(* IEC 61131-3 sources: daoli-st-library/DL_Motion (part 12) *)

(* ---- FB_DL_EdgeTrimTraverse.st ---- *)
(*==============================================================================
 * 组件名称 (Component)  : FB_DL_EdgeTrimTraverse
 * 所属子库 (Sublibrary) : DL_Motion
 * 当前版本 (Version)    : 1.0.0
 * 兼容性 (Platform)     : CODESYS 3.5 / TwinCAT 3 / 汇川 InoProShop（纯标准元素，零方言）
 * 功能描述 (Function)   : 修边刀架横动往复定位。启动后在行程两端之间往复，折返点按重叠量
 *                         外延，端点驻留可组态；停止请求只在段终点生效（半途硬切会在膜面
 *                         留刀痕）。行程过窄、速度出域判组态故障；目标越软包络在启动沿前
 *                         预检拒绝，一轴不动。不做刀压控制、不做随线速度联动、不做多段
 *                         变速。说明：既有 FB_DL_SoftLimitGuard 的契约绑定运动轴接口，
 *                         与本件的开环步进契约不同，故按同一语义内联预检，不做跨契约强转。
 * 溯源 (Origin)         : 道莅 clean-room 防御性实现
 * 本文件内含 (Contains) : TYPE E_DL_TraverseState / FUNCTION_BLOCK FB_DL_EdgeTrimTraverse
 * 依赖 (Depends)        : DL_Device/I_DL_StepperOpenLoop（只调用契约方法与属性）
 * 红线自检 (Redline)    : 无外部全局变量、无硬件地址直引 ｜ 全变量中英双语同行注释
 *                         行程宽度判零防除零 ｜ 重叠量与驻留出域双向钳制 ｜ 非有限用自反比较
 *                         驻留定时器与沿实例无条件周期刷新 ｜ 枚举显式赋值 ｜ CASE 含 ELSE
 * 错误码表 (Codes)      : 16#0004_033B 就绪（空闲/本拍无事件）
 *                         16#0004_033C 故障级 旋转轴/横动轴拒绝运动指令
 *                         16#0004_033D 故障级 组态非法（行程宽度 < 5 mm 或速度出域）
 *                         16#0004_033E 故障级 目标越软包络，启动沿前预检拒绝（一轴不动）
 *                         16#0004_033F 预留：本版不发码（下一轮区间起点，禁止回填）
 * 修订历史 (Revision)   : 2026-11-17  v1.0.0  首版入库 · R28 · 阶段三批 2
 * 验收向量 (Acceptance) : 正向 行程 0~300 mm、100 mm/s、重叠 5 mm、驻留 200 ms → 单程
 *                         约 3 s、端点重叠 5 mm、单程计数 +1
 *                         反向 行程改 0~3 mm（宽 3 mm < 5 mm）→ 16#0004_033D；重叠给
 *                         -50 mm → 钳 0 后照常运行；目标包络外延后越限 → 16#0004_033E
 *                         且一轴不动；轴拒绝指令 → 16#0004_033C
 *============================================================================*)

(*-----------------------------------------------------------------------------
 * 枚举: E_DL_TraverseState（归属本功能块，同文件发布，全库唯一定义）
 * 含义: 横动往复相位，每个成员在 CASE 中有且仅有一个标签。
 *----------------------------------------------------------------------------*)
TYPE E_DL_TraverseState :
(
    eIdle    := 0,    // 空闲：等启动沿与预检 / Idle, waiting for the start edge and the pre-check
    eRunMin  := 10,   // 向负端行进 / Travelling toward the minimum end
    eRunMax  := 20,   // 向正端行进 / Travelling toward the maximum end
    eDwell   := 30,   // 端点驻留计时 / Dwell timing at an end
    eStopped := 40,   // 段终点已停：等停止请求撤除 / Stopped at the segment end, waiting for the stop request to clear
    eFault   := 99    // 故障：锁存码保持，仅启动沿重启 / Fault, the latch code is held until a start edge
);
END_TYPE

FUNCTION_BLOCK FB_DL_EdgeTrimTraverse
VAR_INPUT
    bEnable       : BOOL := FALSE;        // 使能 / Enable
    bStart        : BOOL := FALSE;        // 启动，上升沿启动一次 / Start, the rising edge starts one cycle
    bStop         : BOOL := FALSE;        // 停止，电平请求，段终点生效 / Stop request, level input, effective at the segment end
    fPosMin_mm    : REAL := 0.0;          // 行程负端 [mm]，域 ±1000 / Negative travel end in millimetres, domain plus minus 1000
    fPosMax_mm    : REAL := 300.0;        // 行程正端 [mm]，须 Max − Min ≥ 5 / Positive travel end in millimetres, Max minus Min must reach 5
    fSpeed_mmS    : REAL := 100.0;        // 运行速度 [mm/s]，域 0.5~200 / Run speed in millimetres per second, domain 0.5 to 200
    fOverlap_mm   : REAL := 5.0;          // 端点重叠 [mm]，域 0~20 / End overlap in millimetres, domain 0 to 20
    tDwell        : TIME := T#200MS;      // 端点驻留 [ms]，域 0~5 s / End dwell, domain 0 to 5 s
END_VAR
VAR_IN_OUT
    iAxis         : I_DL_StepperOpenLoop; // 横动轴开环步进契约引用 [—] / Traverse axis open-loop stepper contract reference
END_VAR
VAR_OUTPUT
    fPosOut_mm    : REAL;                 // 当前横动位置 [mm] / Current traverse position in millimetres
    bAtMin        : BOOL;                 // 负端到位 / At the minimum end
    bAtMax        : BOOL;                 // 正端到位 / At the maximum end
    uTraverseCnt  : UDINT;                // 累计单程数 [次] / Accumulated single passes
    eState        : E_DL_TraverseState;   // 横动相位 [—] / Traverse phase
    eErr          : UDINT;                // 错误码，段位 16#0004_xxxx / Error code in segment 16#0004_xxxx
END_VAR
VAR
    _eState       : E_DL_TraverseState := E_DL_TraverseState.eIdle; // 当前相位 / Current phase
    _bInit        : BOOL := FALSE;        // 首扫标志，取非判定 / First-scan flag, tested negated
    _bRefOk       : BOOL;                 // 契约引用有效标志 / Contract reference valid flag
    _bCfgOk       : BOOL;                 // 组态合法标志 / Configuration valid flag
    _bIssueScan   : BOOL;                 // 派单当拍标志（本拍不判就绪） / Dispatch scan flag, readiness is not judged in this scan
    _bStopPending : BOOL;                 // 段终点停止挂起标志 / Stop pending at the segment end
    _bDirMax      : BOOL;                 // 下一段方向：TRUE = 向正端 / Next segment direction, TRUE for the positive end
    _bFaultLatch  : BOOL;                 // 故障锁存标志 / Fault latch flag
    _uLatchCode   : UDINT;                // 锁存码载体 / Latch code carrier
    _fTgtHigh     : REAL;                 // 正端折返目标（含重叠）[mm] / Positive turn target including overlap
    _fTgtLow      : REAL;                 // 负端折返目标（含重叠）[mm] / Negative turn target including overlap
    _fOverlapEff  : REAL := 0.0;          // 生效重叠量（钳制后）[mm] / Effective overlap after clamping
    _fSpeedEff    : REAL := 100.0;        // 生效速度（下限兜底）[mm/s] / Effective speed with a lower bound guard
    _fDist        : REAL;                 // 本段待走距离 [mm] / Pending distance of this segment
    _rtrigStart   : R_TRIG;               // 启动上升沿 / Rising edge of the start command
    _tonDwell     : TON;                  // 端点驻留计时 / End dwell timer
END_VAR
VAR CONSTANT
    DL_TRV_READY   : UDINT := 16#0004_033B;  // 就绪码 / Ready code
    DL_TRV_AXIS_BAD : UDINT := 16#0004_033C; // 故障级轴拒绝码 / Fault code for a rejected axis command
    DL_TRV_CFG_BAD : UDINT := 16#0004_033D;  // 故障级组态非法码 / Fault code for bad configuration
    DL_TRV_LIMIT   : UDINT := 16#0004_033E;  // 故障级预检拒绝码 / Fault code for a pre-check rejection
    DL_TRV_W_MIN   : REAL := 5.0;            // 行程最小宽度 [mm] / Minimum travel width in millimetres
    DL_TRV_POS_HI  : REAL := 1000.0;         // 行程端点绝对值上限 [mm] / Absolute bound of the travel ends
    DL_TRV_OVL_HI  : REAL := 20.0;           // 重叠量上限 [mm] / Overlap upper bound
    DL_TRV_SPD_LO  : REAL := 0.5;            // 速度下限 [mm/s] / Speed lower bound
    DL_TRV_SPD_HI  : REAL := 200.0;          // 速度上限 [mm/s] / Speed upper bound
    DL_TRV_AT_TOL  : REAL := 0.05;           // 端点到位容差 [mm] / End-point arrival tolerance
END_VAR

// 段 1｜输出与单拍标志预置
bAtMin := FALSE;                                    // 负端到位预清 / At-minimum flag pre-cleared
bAtMax := FALSE;                                    // 正端到位预清 / At-maximum flag pre-cleared
eErr := 0;                                          // 错误码预清 / Error code pre-cleared
_bIssueScan := FALSE;                               // 派单当拍标志预清 / Dispatch scan flag pre-cleared

// 段 2｜沿检测无条件周期刷新
_rtrigStart(CLK := bStart);                         // 启动沿 / Start edge

// 段 3｜驻留定时器无条件周期刷新（仅驻留相计时）
_tonDwell(IN := (_eState = E_DL_TraverseState.eDwell), PT := tDwell);

// 段 4｜首扫初始化（判据取非，R19）
IF NOT _bInit THEN
    _eState := E_DL_TraverseState.eIdle;            // 相位待机起步 / Phase starts idle
    _bInit := TRUE;                                 // 首扫只做一次 / The first scan runs once
END_IF

// 段 5｜引用与组态闸（行程宽度 < 5 mm 使往复退化为抖动）
_bRefOk := (iAxis <> 0);
_bCfgOk := _bRefOk
        AND NOT ((fPosMin_mm <> fPosMin_mm) OR ((fPosMin_mm - fPosMin_mm) <> (fPosMin_mm - fPosMin_mm)))
        AND NOT ((fPosMax_mm <> fPosMax_mm) OR ((fPosMax_mm - fPosMax_mm) <> (fPosMax_mm - fPosMax_mm)))
        AND ((fPosMax_mm - fPosMin_mm) >= DL_TRV_W_MIN)
        AND (ABS(fPosMin_mm) <= DL_TRV_POS_HI) AND (ABS(fPosMax_mm) <= DL_TRV_POS_HI)
        AND NOT ((fSpeed_mmS <> fSpeed_mmS) OR ((fSpeed_mmS - fSpeed_mmS) <> (fSpeed_mmS - fSpeed_mmS)))
        AND (fSpeed_mmS >= DL_TRV_SPD_LO) AND (fSpeed_mmS <= DL_TRV_SPD_HI)
        AND (tDwell >= T#0MS) AND (tDwell <= T#5S);
_fSpeedEff := LIMIT(DL_TRV_SPD_LO, fSpeed_mmS, DL_TRV_SPD_HI);          // 生效速度钳制 [mm/s] / Effective speed after clamping
_fOverlapEff := LIMIT(0.0, fOverlap_mm, DL_TRV_OVL_HI);                 // 重叠量钳制 [mm] / Overlap after clamping
_fTgtHigh := fPosMax_mm + _fOverlapEff;                                 // 正端折返目标（外延）[mm] / Positive turn target, extended
_fTgtLow := fPosMin_mm - _fOverlapEff;                                  // 负端折返目标（外延）[mm] / Negative turn target, extended

// 段 6｜位置回读与端点判据
IF _bRefOk THEN
    fPosOut_mm := iAxis.fPosition;                  // 当前横动位置 [mm] / Current traverse position
    bAtMax := ABS(fPosOut_mm - fTgtHigh) <= DL_TRV_AT_TOL;   // 正端到位判据 / At the positive end
    bAtMin := ABS(fPosOut_mm - fTgtLow) <= DL_TRV_AT_TOL;    // 负端到位判据 / At the negative end
ELSE
    fPosOut_mm := 0.0;                              // 引用无效：位置输出置 0 / Invalid reference, the position output is zeroed
END_IF

// 段 7｜失能闸
IF NOT bEnable THEN
    IF _bRefOk THEN
        iAxis.Stop();                               // 失能即受控停车 / Controlled stop on disable
    END_IF
    _eState := E_DL_TraverseState.eIdle;            // 相位回空闲 / Phase back to idle
    _bStopPending := FALSE;                         // 停止挂起清 / Stop pending cleared
    eErr := DL_TRV_READY;                           // 失能为正常停机 / Disable is a normal stop
END_IF

// 段 8｜横动往复状态机（ENUM + CASE + ELSE 兜底）
IF bEnable THEN
    CASE _eState OF

        E_DL_TraverseState.eIdle:                   // 空闲：等启动沿，先做组态与包络预检
            IF _rtrigStart.Q THEN
                _bFaultLatch := FALSE;              // 启动沿为锁存解除路径 / The start edge releases the latch
                _uLatchCode := 0;                   // 锁存码清 / Latch code cleared
                _bStopPending := FALSE;             // 停止挂起清 / Stop pending cleared
                IF NOT _bCfgOk THEN
                    eErr := DL_TRV_CFG_BAD;         // 故障级：组态非法 / Fault, bad configuration
                    _uLatchCode := DL_TRV_CFG_BAD;
                    _bFaultLatch := TRUE;
                    _eState := E_DL_TraverseState.eFault;
                ELSIF (ABS(_fTgtHigh) > DL_TRV_POS_HI) OR (ABS(_fTgtLow) > DL_TRV_POS_HI) THEN
                    eErr := DL_TRV_LIMIT;           // 故障级：重叠外延后越软包络，一轴不动 / Fault, the extended target leaves the envelope
                    _uLatchCode := DL_TRV_LIMIT;
                    _bFaultLatch := TRUE;
                    _eState := E_DL_TraverseState.eFault;
                ELSE
                    _bDirMax := TRUE;               // 首段向正端 / The first segment heads to the positive end
                    _eState := E_DL_TraverseState.eRunMax;
                END_IF
            ELSE
                IF NOT _bCfgOk THEN
                    eErr := DL_TRV_CFG_BAD;         // 故障级：组态非法（空闲期即报） / Fault, bad configuration reported while idle
                    _uLatchCode := DL_TRV_CFG_BAD;
                    _bFaultLatch := TRUE;
                    _eState := E_DL_TraverseState.eFault;
                END_IF
            END_IF

        E_DL_TraverseState.eRunMax:                 // 向正端行进：等轴就绪，停止请求挂起
            IF _bIssueScan THEN
                _bIssueScan := FALSE;               // 派单拍已过 / The dispatch scan has passed
            ELSIF (NOT _bStopPending) AND bStop THEN
                _bStopPending := TRUE;              // 停止请求挂起，段终点生效 / Stop pending, effective at the segment end
            ELSIF iAxis.bReady THEN
                uTraverseCnt := uTraverseCnt + 1;   // 单程计数 +1 [次] / Single-pass count incremented
                IF _bStopPending THEN
                    _eState := E_DL_TraverseState.eStopped;   // 段终点停车 / Stop at the segment end
                ELSE
                    _eState := E_DL_TraverseState.eDwell;     // 端点驻留 / Dwell at the end
                END_IF
            END_IF

        E_DL_TraverseState.eRunMin:                 // 向负端行进：等轴就绪，停止请求挂起
            IF _bIssueScan THEN
                _bIssueScan := FALSE;
            ELSIF (NOT _bStopPending) AND bStop THEN
                _bStopPending := TRUE;
            ELSIF iAxis.bReady THEN
                uTraverseCnt := uTraverseCnt + 1;   // 单程计数 +1 [次] / Single-pass count incremented
                IF _bStopPending THEN
                    _eState := E_DL_TraverseState.eStopped;
                ELSE
                    _eState := E_DL_TraverseState.eDwell;
                END_IF
            END_IF

        E_DL_TraverseState.eDwell:                  // 端点驻留：计时满后换向派单
            IF _tonDwell.Q THEN
                IF _bDirMax THEN
                    _bDirMax := FALSE;              // 换向：下一段向负端 / Reverse, the next segment heads to the negative end
                    _fDist := _fTgtLow - iAxis.fPosition;      // 待走距离 [mm] / Pending distance
                ELSE
                    _bDirMax := TRUE;               // 换向：下一段向正端 / Reverse, the next segment heads to the positive end
                    _fDist := _fTgtHigh - iAxis.fPosition;     // 待走距离 [mm] / Pending distance
                END_IF
                IF iAxis.MoveRelative(_fDist, _fSpeedEff) THEN
                    _bIssueScan := TRUE;            // 派单当拍不判就绪 / Readiness is not judged in the dispatch scan
                    IF _bDirMax THEN
                        _eState := E_DL_TraverseState.eRunMax;
                    ELSE
                        _eState := E_DL_TraverseState.eRunMin;
                    END_IF
                    eErr := DL_TRV_READY;           // 就绪码 / Ready code
                ELSE
                    eErr := DL_TRV_AXIS_BAD;        // 故障级：轴拒绝指令 / Fault, the axis rejected the command
                    _uLatchCode := DL_TRV_AXIS_BAD;
                    _bFaultLatch := TRUE;
                    _eState := E_DL_TraverseState.eFault;
                END_IF
            END_IF

        E_DL_TraverseState.eStopped:                // 段终点已停：停止请求撤除后回空闲
            IF NOT bStop THEN
                _bStopPending := FALSE;
                _eState := E_DL_TraverseState.eIdle;
            END_IF
            eErr := DL_TRV_READY;

        E_DL_TraverseState.eFault:                  // 故障：锁存码保持，仅新启动沿重启
            eErr := _uLatchCode;                    // 锁存码回放 / Replay the latch code
            IF _rtrigStart.Q THEN
                _bFaultLatch := FALSE;
                _uLatchCode := 0;
                _bStopPending := FALSE;
                eErr := DL_TRV_READY;
                _eState := E_DL_TraverseState.eIdle; // 回空闲需再给启动沿（下一拍） / A further start edge is required
            END_IF

        ELSE
            // 非法状态兜底（故障级）
            eErr := DL_TRV_CFG_BAD;                 // 故障级：非法相位 / Fault, illegal phase
            _uLatchCode := DL_TRV_CFG_BAD;
            _bFaultLatch := TRUE;
            _eState := E_DL_TraverseState.eFault;

    END_CASE
END_IF

eState := _eState;                                  // 相位出口镜像 / Phase mirrored to the output pin
END_FUNCTION_BLOCK

(* ---- FB_DL_ElectrodeRollDiameter.st ---- *)
// =====================================================================
// FB_DL_ElectrodeRollDiameter.st
// 极卷直径跟踪与换卷预警（卷径递推 + 低速保护 + 单调校核 + 换卷阈值预警）
// Electrode roll diameter tracking with change-over warning
// 所属子库: DL_Motion    版本: v1.0.0    兼容: CODESYS V3.5+ / TwinCAT 3 / 汇川 InoProShop
// 码位: 16#0004_035E ~ 16#0004_0362 (本件独占 5 槽, 勿复用)
// 溯源: 道莅 clean-room 防御性实现
//       来源组标签: lithium-battery, winding, coil-diameter, warning
// 修改记录: R30 初版 (ROUND_PLAN_R30 序 16)
// 分层声明: 卷径换算公式与 FC_DL_CoilDiameterCalc 口径一致（本件只加跟踪
//           与预警层, 不重写公式件）: D = v·k/(π·n), k = 1000 mm/m
// =====================================================================
FUNCTION_BLOCK FB_DL_ElectrodeRollDiameter
VAR_INPUT
    fLineSpd_mmin : REAL := 0.0;    // 线速度 0~300 m/min / Line speed [m/min]
    fRollRpm      : REAL := 0.0;    // 卷轴转速 0~3000 r/min / Roll speed [r/min]
    fPrevDia_mm   : REAL := 500.0;  // 上次卷径注入 0~2000 mm / Previous diameter injected [mm]
    fCoreDia_mm   : REAL := 76.0;   // 卷芯直径 0~2000 mm / Core diameter [mm]
    fThick_um     : REAL := 25.0;   // 层厚校核值 0~500 um / Layer thickness [um]
    fWarnDia_mm   : REAL := 120.0;  // 换卷预警径 0~2000 mm / Change warning diameter [mm]
END_VAR
VAR_OUTPUT
    fDia_mm     : REAL := 0.0;      // 当前卷径 / Current diameter [mm]
    bChangeWarn : BOOL := FALSE;    // 换卷预警 / Change-over warning
    bAtCore     : BOOL := FALSE;    // 卷径触及芯径 / At core flag
    eErr        : UDINT := 16#0004_035E;  // 错误码 / Error code
END_VAR
VAR
    rPi     : REAL := 3.14159265358979;   // 圆周率 / Pi constant
    fSpdMin : REAL := 1.0;          // 低速门限（线速度）m/min, 工程固定门限 / Min line speed gate
    fRpmMin : REAL := 5.0;          // 低速门限（转速）r/min, 工程固定门限 / Min roll speed gate
    fCalcDia: REAL := 0.0;          // 本拍换算卷径 / Calculated diameter this cycle [mm]
    fTolDia : REAL := 0.0;          // 单调校核容差（双倍层厚换算）/ Monotonic tolerance from thickness [mm]
    bCfgErr : BOOL := FALSE;        // 组态非法标记 / Configuration error flag
    bHoldErr: BOOL := FALSE;        // 递推保持标记（非有限或单调违反）/ Recursion hold flag
    bLowSpd : BOOL := FALSE;        // 低速保护标记 / Low speed protection flag
    xFirst  : BOOL := TRUE;         // 首扫标记 / First-scan flag
END_VAR

// ---------------------------------------------------------------------
// 代码位表（本件独占, 勿复用）:
//   16#0004_035E 信息 卷径跟踪正常
//   16#0004_035F 故障 组态非法（芯径/预警径非有限或不大于 0, 或芯径不低于
//                预警径倒置）; 解除式 = 恢复合法组态
//   16#0004_0360 故障 递推保持（速度/转速非有限, 或新卷径违反放卷单调递减）,
//                卷径保持上拍值; 解除式 = 输入恢复有限且差分恢复单调
//   16#0004_0361 信息 低速保护冻结（线速或转速低于门限, 卷径保持不递推）
//   16#0004_0362 信息 换卷预警（卷径不大于预警径, 含触及芯径）
// ---------------------------------------------------------------------

// ---- 首扫: 以注入的上次卷径为初始跟踪值 / First scan: seed from injected ----
IF xFirst THEN
    fDia_mm := fPrevDia_mm;     // 初始卷径 / Initial diameter [mm]
    xFirst := FALSE;            // 清首扫标记 / Clear flag
END_IF

// ---- 组态闸 / Configuration gate ----
bCfgErr := FALSE;
IF (fCoreDia_mm <> fCoreDia_mm) OR (fCoreDia_mm <= 0.0) OR (fCoreDia_mm > 2000.0) THEN
    bCfgErr := TRUE;            // 芯径非法 / Illegal core diameter
END_IF
IF (fWarnDia_mm <> fWarnDia_mm) OR (fWarnDia_mm <= 0.0) OR (fWarnDia_mm > 2000.0) THEN
    bCfgErr := TRUE;            // 预警径非法 / Illegal warning diameter
END_IF
IF (NOT bCfgErr) AND (fCoreDia_mm >= fWarnDia_mm) THEN
    bCfgErr := TRUE;            // 芯径不低于预警径 = 倒置 / Inverted config
END_IF

// ---- 输出缺省 / Output defaults ----
bHoldErr := FALSE;
bLowSpd  := FALSE;

IF bCfgErr THEN
    // 组态非法: 卷径保持, 安全侧不递推 / Config fault: hold, no recursion
    eErr := 16#0004_035F;
ELSE
    // ---- 低速保护判 / Low speed protection judge ----
    bLowSpd := (fLineSpd_mmin < fSpdMin) OR (fRollRpm < fRpmMin);
    // ---- 非有限判 / Finite judge ----
    IF (fLineSpd_mmin <> fLineSpd_mmin) OR (ABS(fLineSpd_mmin) >= 1.0E12)
       OR (fRollRpm <> fRollRpm) OR (ABS(fRollRpm) >= 1.0E12)
       OR (fPrevDia_mm <> fPrevDia_mm) THEN
        bHoldErr := TRUE;       // 非有限保持 / Non-finite hold
        eErr := 16#0004_0360;
    ELSIF bLowSpd THEN
        // 低速保护: 冻结递推, 卷径保持 / Freeze recursion on low speed
        eErr := 16#0004_0361;
    ELSE
        // ---- 卷径递推: D = v·k/(π·n), k = 1000 mm/m, 转速门限已保证不为零
        //      Diameter recursion with guarded division ----
        fCalcDia := (fLineSpd_mmin * 1000.0) / (rPi * fRollRpm);
        // 层厚校核容差: 允许的单拍回升量 = 两倍层厚换算 / Monotonic tolerance from thickness
        fTolDia := 2.0 * fThick_um / 1000.0;
        IF fCalcDia > (fDia_mm + fTolDia) THEN
            // 放卷单调递减违反: 保持 + 故障码 / Monotonic violation: hold
            bHoldErr := TRUE;
            eErr := 16#0004_0360;
        ELSE
            fDia_mm := fCalcDia;    // 递推更新 / Update diameter
            // 卷径下限钳卷芯径 / Clamp to core diameter
            IF fDia_mm < fCoreDia_mm THEN
                fDia_mm := fCoreDia_mm;
            END_IF
            eErr := 16#0004_035E;   // 跟踪正常 / Tracking normal
        END_IF
    END_IF
END_IF

// ---- 预警与触芯输出（闭口径: 恰好等于预警径即触发）/ Warning and at-core ----
bChangeWarn := fDia_mm <= fWarnDia_mm;      // 恰好等于预警径与更低均触发 / Trigger at and below
bAtCore := (fDia_mm - fCoreDia_mm) < 1.0E-6;    // 容差判触芯 / At core with tolerance

END_FUNCTION_BLOCK

(* ---- FB_DL_ElectronicCamSwitchBank.st ---- *)
(*
  FB_DL_ElectronicCamSwitchBank  —  电子凸轮开关组（MC_CamSwitch 语义）/ Electronic cam switch bank
  分类 Category : DL_Motion
  码位 Code     : 16#04_0_A5
  版本 Version  : 1.0.0
  来源 Source   : t1-6-plcopen — IEC 61131-3 标准语义的道莅防御性实现
  溯源 Origin   : PLCopen MC_CamSwitch 公开语义借鉴，clean-room 实现，未复制任何源码行
                  （与 FB_DL_MarkPositionLatch 分工相反：本件由位置产生输出；FB_DL_ElectronicCam 管凸轮表插值，本件只做开关窗判）
  功能 Function : 1) 轴位置（模 360）逐路判是否落在 [pos+offset, pos+offset+width]；窗口跨 0° 按两段拆判；
                  2) Cyclic 每圈重复触发；Single 每开关只触发一次（abFired 锁存，重置仅经 bReset 上升沿）；
                  3) nActiveMask 聚合 ≤32 路活动位（SHL 显式位号，禁魔法掩码）。
  边界 Boundary : ① uSwitchCount = 0 或超数组上界（32）判组态错返回（全输出 FALSE 安全侧）；
                  ② uSwitchCount > 32 不生成 nActiveMask（判组态错，禁静默截断）；
                  ③ afSwitchWidthDeg <= 0 或 >= 360 判组态错；
                  ④ 轴位置非有限（NaN 用 x<>x 自反判定）置故障态并全输出 FALSE（安全侧，锁存至复位）；
                  ⑤ 解除式自证：abFired 清零 = bReset 上升沿（引脚可满足）；Fault 退出 = bReset 上升沿 AND 组态合法；
                  ⑥ CASE 全态覆盖 + ELSE 兜底置故障相。
  依赖 Depends  : I_DL_MotionAxis（注入，不实例化）；仅 Standard.library（R_TRIG/SHL）
  码表 Error codes（本件格 04_0_A5，子码步进 +0x100）:
    16#0004_01A5 信息级：开关组使能运行中（不置故障）
    16#0004_02A5 故障级：组态非法（通道数越域 / 宽度 <= 0 或 >= 360），锁存至复位
    16#0004_03A5 故障级：轴位置非有限（NaN/Inf），全输出 FALSE，锁存至复位
    16#0004_04A5 故障级：状态机落 ELSE 兜底（非法相位 ID）

  修订历史 Revision :
    2026-11-18  v1.0.0  R38 首版
*)

TYPE E_DL_CamSwMode :
(
    eSingle := 0,   // 单次：每开关每使能期只触发一次 / Single, fires once per enable period
    eCyclic := 1    // 周期：每圈重复触发 / Cyclic, fires every revolution
);
END_TYPE

TYPE E_DL_CamSwState :
(
    eIdle  := 0,    // 空闲：未使能 / Idle, not enabled
    eRun   := 10,   // 运行：使能且位置有效 / Run, enabled with valid position
    eFault := 90    // 故障：组态/位置故障锁定 / Fault, latched
);
END_TYPE

FUNCTION_BLOCK FB_DL_ElectronicCamSwitchBank
VAR_INPUT
    anSwitchPosDeg  : ARRAY[0..31] OF LREAL;   // 开关位置表 [deg] / Switch position table
    afSwitchWidthDeg: ARRAY[0..31] OF REAL;    // 触发宽度 [deg] / Trigger width
    auPhaseOffsetDeg: ARRAY[0..31] OF REAL;    // 相位偏移 [deg] / Phase offset
    uSwitchCount    : INT;                     // 开关数 [路]，域 1..32 / Switch count
    bEnable         : BOOL := FALSE;           // 使能 / Enable
    eTriggerMode    : E_DL_CamSwMode;          // 触发模式（Single/Cyclic）/ Trigger mode
    bReset          : BOOL := FALSE;           // 复位（abFired 清零唯一路径）/ Reset, sole abFired clear path
END_VAR
VAR_OUTPUT
    abSwitchOut     : ARRAY[0..31] OF BOOL;    // 各开关输出 / Per-switch outputs
    bAnyActive      : BOOL;                    // 任一开关活动 / Any switch active
    nActiveMask     : DWORD;                   // 活动位掩码（<= 32 路才生成）/ Active bit mask
    nErrId          : UDINT;                   // 事件码，0 = 无事件 / Event code
    eState          : E_DL_CamSwState;         // 状态出口，段尾单点映射 / State outlet
END_VAR
VAR_IN_OUT
    iAxis           : I_DL_MotionAxis;         // 轴接口引用（注入，不实例化）/ Axis reference, injected
END_VAR
VAR
    rtReset  : R_TRIG;                         // 复位上升沿 / Reset rising edge
    _eState  : E_DL_CamSwState := E_DL_CamSwState.eIdle;   // 内部相位（CASE 唯一写入目标）/ Internal phase
    _abFired : ARRAY[0..31] OF BOOL;           // Single 模式已触发锁存 / Single-mode fired latch
    _bCfgBad : BOOL;                           // 组态非法锁存 / Configuration fault latch
    _bPosBad : BOOL;                           // 位置非有限标志 / Position non-finite flag
    _rPos    : LREAL;                          // 轴位置 [deg] / Axis position
    _rPosMod : LREAL;                          // 模 360 位置 [deg] / Position modulo 360
    _rStart  : LREAL;                          // 窗口起点（模 360）/ Window start, wrapped
    _rEnd    : LREAL;                          // 窗口终点（模 360 前）/ Window end before wrap
    _bInWin  : BOOL;                           // 本路在窗标志 / In-window flag
    _nK      : INT;                            // 循环计数器 / Loop counter
END_VAR
VAR CONSTANT
    nMaxSw     : INT   := 32;      // 数组上界 = 掩码位宽 [路] / Array bound = mask width
    DL_FULL    : LREAL := 360.0;   // 全圆周期 [deg] / Full circle period
    DL_ZERO_EPS: LREAL := 1.0E-9;  // 近零判据 / Near-zero epsilon
END_VAR

(* —— 段 0：边沿无条件周期刷新（R182：调用语句不得置于 IF/CASE 内） —— *)
rtReset(CLK := bReset);                        // 复位上升沿，每拍必调

(* —— 段 1：单拍量预清零（锁存量 _abFired/_bCfgBad 不入清单，R187①） —— *)
bAnyActive := FALSE;                           // 聚合出口缺省 FALSE
nActiveMask := 0;                              // 掩码缺省 0
nErrId := 16#0000_0000;                        // 事件码缺省无事件
FOR _nK := 0 TO (nMaxSw - 1) DO
    abSwitchOut[_nK] := FALSE;                 // 输出缺省 FALSE（安全侧，段 6 单点置位）
END_FOR

(* —— 段 2：复位沿（abFired 清零唯一路径；Fault 解除唯一路径） —— *)
IF rtReset.Q THEN
    FOR _nK := 0 TO (nMaxSw - 1) DO
        _abFired[_nK] := FALSE;                // Single 触发锁存清零（解除式自证：bReset 可满足）
    END_FOR
    _bCfgBad := FALSE;                         // 组态锁存清零
    _bPosBad := FALSE;                         // 位置故障清零
    IF _eState = E_DL_CamSwState.eFault THEN
        _eState := E_DL_CamSwState.eIdle;      // 故障相回空闲（组态合法性由段 3 复判）
    END_IF
END_IF

(* —— 段 3：组态域闸（每拍复判；锁存置位只在 Fault 判定时引用） —— *)
IF (uSwitchCount <= 0) OR (uSwitchCount > nMaxSw) THEN
    _bCfgBad := TRUE;                          // 通道数越域（> 32 不生成掩码，禁静默截断）
END_IF
IF NOT _bCfgBad THEN
    FOR _nK := 0 TO (uSwitchCount - 1) DO
        IF (LREAL(afSwitchWidthDeg[_nK]) <= DL_ZERO_EPS)
           OR (LREAL(afSwitchWidthDeg[_nK]) >= DL_FULL) THEN
            _bCfgBad := TRUE;                  // 宽度 <= 0 或 >= 360
        END_IF
        IF (REAL_TO_LREAL(auPhaseOffsetDeg[_nK]) <> REAL_TO_LREAL(auPhaseOffsetDeg[_nK]))
           OR (ABS(REAL_TO_LREAL(auPhaseOffsetDeg[_nK])) >= DL_FULL) THEN
            _bCfgBad := TRUE;                  // 相位偏移非有限或越一圈
        END_IF
    END_FOR
END_IF

(* —— 段 4：轴位置采集与非有限判定（NaN 用 x<>x 自反，Inf 用幅值上限兜） —— *)
_rPos := iAxis.fPosition;                      // 轴位置 [deg]
IF (_rPos <> _rPos) OR (ABS(_rPos) > 1.0E15) THEN
    _bPosBad := TRUE;                          // 非有限：置故障态全输出 FALSE（安全侧）
END_IF
IF NOT _bPosBad THEN
    _rPosMod := _rPos - DL_FULL * TRUNC(_rPos / DL_FULL);   // 模 360 折返到 [0, 360)
END_IF

(* —— 段 5：相位机（只做迁移；出口在段 6） —— *)
CASE _eState OF

E_DL_CamSwState.eIdle:
    IF _bCfgBad OR _bPosBad THEN
        _eState := E_DL_CamSwState.eFault;     // 组态/位置故障：进故障相
    ELSIF bEnable THEN
        _eState := E_DL_CamSwState.eRun;       // 使能：进运行相
    END_IF

E_DL_CamSwState.eRun:
    IF _bCfgBad OR _bPosBad THEN
        _eState := E_DL_CamSwState.eFault;     // 组态/位置故障：进故障相
    ELSIF NOT bEnable THEN
        _eState := E_DL_CamSwState.eIdle;      // 失能：回空闲（故障与失能分流，归因唯一）
    END_IF

E_DL_CamSwState.eFault:
    ;                                          // 故障相：等复位沿（段 2 承载解除）

ELSE
    _eState := E_DL_CamSwState.eFault;         // 非法相位 ID 兜底

END_CASE

(* —— 段 6：窗口判算与出口（仅运行相执行；故障/空闲全 FALSE 已由段 1 缺省保证） —— *)
IF _eState = E_DL_CamSwState.eRun THEN
    FOR _nK := 0 TO (uSwitchCount - 1) DO
        _rStart := _rPosMod + LREAL(auPhaseOffsetDeg[_nK]);     // 起点 = 位置 + 相位偏移
        _rStart := _rStart - DL_FULL * TRUNC(_rStart / DL_FULL); // 模 360 折返到 [0, 360)
        _rEnd   := _rStart + LREAL(afSwitchWidthDeg[_nK]);      // 终点（可越 360）
        IF _rEnd <= DL_FULL THEN
            _bInWin := (_rPosMod >= _rStart) AND (_rPosMod <= _rEnd);            // 单段判
        ELSE
            _bInWin := (_rPosMod >= _rStart) OR (_rPosMod <= (_rEnd - DL_FULL)); // 跨 0° 两段拆判
        END_IF
        IF _bInWin THEN
            IF eTriggerMode = E_DL_CamSwMode.eSingle THEN
                IF NOT _abFired[_nK] THEN
                    abSwitchOut[_nK] := TRUE;       // Single：首遇触发
                    _abFired[_nK] := TRUE;          // 触发锁存（bReset 沿清零）
                END_IF
            ELSE
                abSwitchOut[_nK] := TRUE;           // Cyclic：每圈重复触发
            END_IF
            nActiveMask := nActiveMask OR SHL(INT_TO_DWORD(1), _nK);   // SHL 显式位号（禁魔法掩码）
        END_IF
    END_FOR
    bAnyActive := nActiveMask <> 0;                 // 任一活动聚合
    nErrId := 16#0004_01A5;                         // 信息级：开关组运行中
END_IF

(* —— 段 7：故障码与状态出口单点映射（锁存码回放，禁同拍抹除） —— *)
IF (_eState = E_DL_CamSwState.eFault) AND _bCfgBad THEN
    nErrId := 16#0004_02A5;                         // 故障级：组态非法
ELSIF (_eState = E_DL_CamSwState.eFault) AND _bPosBad THEN
    nErrId := 16#0004_03A5;                         // 故障级：位置非有限
END_IF
eState := _eState;                                  // 状态出口单点映射

END_FUNCTION_BLOCK

(* ---- FB_DL_ElectronicLineShaftSeq.st ---- *)
(*
  Name: FB_DL_ElectronicLineShaftSeq
  Category: DL_Motion
  Version: 1.0.0
  Round: R89 / 2026-11-25
  开源溯源：clean-room 自研（族 运动同步控制，ST 开源生态实测 0 命中，无外部代码引入）
  功能：电子线轴多从站同步：主轴相位广播 + 逐从站偏置斜坡 + 使能时序，偏置超限即拒并使能。
  边界条件：① 五浮点入参（主轴转速、偏置上限、周期）与四元素偏置数组全部过非有限闸；
            ② 主轴相位按 rpm × 6 × 周期 累加（1 r/min = 6 °/s），保持 [0,360) 防长时精度流失；
            ③ 逐从站偏置斜坡：目标 = anSlaveOffsetDeg[i]，速率 DL_ELS_RATE [°/s]，步长 = 速率 × fCycleS；
            ④ 偏置绝对值超 fMaxOffsetDeg 即拒绝使能：故障锁存 + 四从站速度给定全部置 0（安全侧）；
            ⑤ 未就绪从站（anSlaveReady = FALSE）不参与同步，nSlaveOnline 照实计数，xAllSynced 必须四站齐备；
            ⑥ 故障解除唯一路径：故障相内 xEnable 释放（R152），清锁存回 eIdle。
  状态机：eIdle / eEnable / eRamp / eSynced / eFault（CASE 含 ELSE 兜底）。
  量纲自证：rpm × 6 = °/s；°/s × s = °；°/s × s = °（偏置步长）。
*)
TYPE E_DL_ElsPhase :
(
    eIdle   := 0,       (* 待机：等使能沿 / Idle, waiting for enable edge *)
    eEnable := 10,      (* 使能相：核从站在线数与偏置上限 / Enable check *)
    eRamp   := 20,      (* 斜坡相：逐从站偏置斜坡 / Offset ramping *)
    eSynced := 30,      (* 同步相：相位广播运行 / Synced, phase broadcast *)
    eFault  := 90       (* 故障相：锁存待释放 / Fault latched, awaiting release *)
);
END_TYPE

FUNCTION_BLOCK FB_DL_ElectronicLineShaftSeq
VAR_INPUT
    xEnable : BOOL;                                 (* 使能 [-] Enable *)
    fMasterVelRpm : REAL;                           (* 主轴速度 [r/min] Master velocity [rpm] *)
    anSlaveOffsetDeg : ARRAY[1..4] OF REAL;         (* 四从站相位偏置目标 [°] Slave phase offsets [deg] *)
    anSlaveReady : ARRAY[1..4] OF BOOL;             (* 四从站就绪反馈 [-] Slave ready feedback *)
    fMaxOffsetDeg : REAL;                           (* 偏置允许上限（绝对值） [°] Offset magnitude limit [deg] *)
    fCycleS : REAL;                                 (* 扫描周期 [s] Scan cycle [s] *)
END_VAR
VAR_OUTPUT
    anSlaveVelRefRpm : ARRAY[1..4] OF REAL;         (* 四从站速度给定 [r/min] Slave velocity references [rpm] *)
    xAllSynced : BOOL;                              (* 四从站全部同步 [-] All slaves synced *)
    nSlaveOnline : INT;                             (* 在线（就绪）从站数 0~4 [站] Online slave count *)
    xFault : BOOL;                                  (* 故障锁存标志 [-] Fault latched *)
END_VAR
VAR
    _eState : E_DL_ElsPhase := E_DL_ElsPhase.eIdle;  (* 内部相（CASE 唯一写入目标） [-] Internal phase *)
    _bInit : BOOL := FALSE;                         (* 首扫初始化标志 [-] First-scan init flag *)
    _bFaultLatch : BOOL := FALSE;                   (* 故障锁存位 [-] Fault latch *)
    _bReqFault : BOOL := FALSE;                     (* 单拍故障请求（段 2 预清） [-] Fault request *)
    _bCfgBad : BOOL := FALSE;                       (* 配置非法当拍量 [-] Configuration bad *)
    _bLimBad : BOOL := FALSE;                       (* 偏置超限当拍量 [-] Offset over limit *)
    _bRampDone : BOOL := FALSE;                     (* 四站偏置斜坡全部到位 [-] All ramps complete *)
    _nOnline : INT := 0;                            (* 就绪计数 [站] Ready count *)
    _nI : INT := 1;                                 (* 从站遍历索引 [-] Slave loop index *)
    _fCy : REAL := 0.01;                            (* 当拍有效周期 [s] Effective cycle [s] *)
    _fMasterPhaseDeg : REAL := 0.0;                 (* 主轴相位保持量 [°] Master phase hold [deg] *)
    _fAdvDeg : REAL := 0.0;                         (* 单拍主轴相位增量 [°] Master phase increment [deg] *)
    _fOffStep : REAL := 0.0;                        (* 单拍偏置斜坡步长 [°] Offset ramp step [deg] *)
    _afOffRamp : ARRAY[1..4] OF REAL;               (* 四从站偏置斜坡当前值 [°] Offset ramp values [deg] *)
    _afVelRef : ARRAY[1..4] OF REAL;                (* 四从站速度给定内部量 [r/min] Velocity ref internal [rpm] *)
    rtEnable : R_TRIG;                              (* 使能沿（段 1 无条件调用） / Enable edge *)
    _bMasterOk : BOOL;                              (* 主轴转速给定有效位（非有限/越限即假） / Master vel valid *)
END_VAR
VAR CONSTANT
    DL_ELS_EPS : REAL := 1.0E-9;        (* 判据容差 [-] Criterion tolerance *)
    DL_ELS_RATE : REAL := 90.0;         (* 偏置斜坡速率 [°/s] Offset ramp rate [deg/s] *)
    DL_ELS_TOL : REAL := 0.5;           (* 偏置到位容差 [°] Offset tolerance [deg] *)
    DL_ELS_CYDEF : REAL := 0.01;        (* 缺省扫描周期 [s] Default scan cycle [s] *)
    DL_ELS_RPM_DEG : REAL := 6.0;       (* 转速 → 角速度换算 [°/s per rpm] Rpm to deg per second *)
    DL_ELS_FULL : REAL := 360.0;        (* 整转角度 [°] Full revolution [deg] *)
    DL_ELS_SNUM : INT := 4;             (* 从站总数 [-] Slave count *)
    DL_ELS_ON_MAX : REAL := 3600.0;     (* 主轴速度上限 [r/min] Master velocity ceiling [rpm] *)
    DL_ELS_OFF_MAX : REAL := 360.0;     (* 偏置上限的工程上限 [°] Offset limit ceiling [deg] *)
END_VAR
(* —— 段 0：非有限闸（NaN 自反 + Inf 差值自减）+ 组态域闸，含四元素偏置数组全枚举（R272） —— *)
_bCfgBad := (fMasterVelRpm <> fMasterVelRpm) OR ((fMasterVelRpm - fMasterVelRpm) <> 0.0)
         OR (fMaxOffsetDeg <> fMaxOffsetDeg) OR ((fMaxOffsetDeg - fMaxOffsetDeg) <> 0.0)
         OR (fCycleS <> fCycleS) OR ((fCycleS - fCycleS) <> 0.0)
         OR (fMasterVelRpm < 0.0) OR (fMasterVelRpm > DL_ELS_ON_MAX)
         OR (fMaxOffsetDeg < 1.0) OR (fMaxOffsetDeg > DL_ELS_OFF_MAX);
FOR _nI := 1 TO DL_ELS_SNUM DO
    IF (anSlaveOffsetDeg[_nI] <> anSlaveOffsetDeg[_nI])
       OR ((anSlaveOffsetDeg[_nI] - anSlaveOffsetDeg[_nI]) <> 0.0) THEN
        _bCfgBad := TRUE;                       (* 偏置数组非有限 / Offset array non-finite *)
    END_IF
END_FOR
(* 周期派生：非法周期取 10 ms 缺省 *)
IF (fCycleS > 0.0) AND (fCycleS <= 1.0) THEN
    _fCy := fCycleS;
ELSE
    _fCy := DL_ELS_CYDEF;
END_IF
(* 主轴相位增量：rpm × 6 = °/s，× s = ° *)
_fAdvDeg := fMasterVelRpm * DL_ELS_RPM_DEG * _fCy;
(* 首扫初始化：偏置斜坡与速度给定归零（R310） *)
IF NOT _bInit THEN
    FOR _nI := 1 TO DL_ELS_SNUM DO
        _afOffRamp[_nI] := 0.0;
        _afVelRef[_nI] := 0.0;
    END_FOR
    _bInit := TRUE;
END_IF
(* —— 段 0：主轴转速有效性单点算定（NOT(x<=lim) 对 NaN 为真 → 判假，防 NaN 直穿速度给定） —— *)
_bMasterOk := (fMasterVelRpm <= 10000.0) AND (fMasterVelRpm >= -10000.0);

(* —— 段 1：偏置斜坡推进 + 超限判定 + 速度给定派生（逐从站，FOR 计数配对） —— *)
_bRampDone := TRUE;
_bLimBad := FALSE;
_fOffStep := DL_ELS_RATE * _fCy;
FOR _nI := 1 TO DL_ELS_SNUM DO
    (* 偏置上限（绝对值）判定：先判目标再判斜坡值 *)
    IF (anSlaveOffsetDeg[_nI] > fMaxOffsetDeg) OR (anSlaveOffsetDeg[_nI] < (0.0 - fMaxOffsetDeg))
       OR (_afOffRamp[_nI] > fMaxOffsetDeg) OR (_afOffRamp[_nI] < (0.0 - fMaxOffsetDeg)) THEN
        _bLimBad := TRUE;                       (* 偏置越限 / Offset over limit *)
    END_IF
    (* 斜坡推进：向目标步进，禁越过目标 *)
    IF _afOffRamp[_nI] < (anSlaveOffsetDeg[_nI] - DL_ELS_TOL) THEN
        _afOffRamp[_nI] := _afOffRamp[_nI] + _fOffStep;
        IF _afOffRamp[_nI] > anSlaveOffsetDeg[_nI] THEN
            _afOffRamp[_nI] := anSlaveOffsetDeg[_nI];
        END_IF
    ELSIF _afOffRamp[_nI] > (anSlaveOffsetDeg[_nI] + DL_ELS_TOL) THEN
        _afOffRamp[_nI] := _afOffRamp[_nI] - _fOffStep;
        IF _afOffRamp[_nI] < anSlaveOffsetDeg[_nI] THEN
            _afOffRamp[_nI] := anSlaveOffsetDeg[_nI];
        END_IF
    END_IF
    IF ABS(_afOffRamp[_nI] - anSlaveOffsetDeg[_nI]) > DL_ELS_TOL THEN
        _bRampDone := FALSE;                    (* 任一未到位即未完成 / Any ramp incomplete *)
    END_IF
    (* 速度给定：使能且未越限且就绪才跟随主轴，否则 0（安全侧） *)
    IF xEnable AND (NOT _bLimBad) AND (NOT _bFaultLatch) AND anSlaveReady[_nI] THEN
        (* 主轴转速非有限/越限闸：NOT(x<=lim) 对 NaN 为真 → 给定归零 *)
        IF _bMasterOk THEN
            _afVelRef[_nI] := fMasterVelRpm;
        ELSE
            _afVelRef[_nI] := 0.0;
        END_IF
        ELSE
        _afVelRef[_nI] := 0.0;                  (* 安全侧：不跟随 / Safe side, no follow *)
    END_IF
END_FOR
(* 就绪计数 *)
_nOnline := 0;
FOR _nI := 1 TO DL_ELS_SNUM DO
    IF anSlaveReady[_nI] THEN
        _nOnline := _nOnline + 1;
    END_IF
END_FOR
(* —— 段 2：单拍量预清 + 故障请求（组态/偏置超限） —— *)
_bReqFault := FALSE;
IF _bCfgBad OR _bLimBad THEN
    _bReqFault := TRUE;                         (* 组态坏或偏置越限：拒并使能 / Rejected *)
END_IF
(* —— 段 3：故障锁存解除（唯一路径 = 故障相内 xEnable 释放，R152） —— *)
IF _bFaultLatch AND (NOT xEnable) THEN
    _bFaultLatch := FALSE;                      (* 清锁存 / Clear latch *)
    _eState := E_DL_ElsPhase.eIdle;             (* 迁回待机 / Back to idle *)
END_IF
(* —— 段 4：使能沿无条件刷新（R7） —— *)
rtEnable(CLK := xEnable);
(* —— 段 5：主状态机（ENUM + CASE，ELSE 兜底） —— *)
CASE _eState OF
E_DL_ElsPhase.eIdle:
    IF rtEnable.Q AND (NOT _bFaultLatch) THEN
        _eState := E_DL_ElsPhase.eEnable;       (* 使能沿 → 使能核查相 / Enable check *)
    END_IF
E_DL_ElsPhase.eEnable:
    IF _nOnline < DL_ELS_SNUM THEN
        _eState := E_DL_ElsPhase.eEnable;       (* 从站未齐：驻留核查（不推进相位） / Wait all ready *)
    ELSIF NOT xEnable THEN
        _eState := E_DL_ElsPhase.eIdle;
    ELSE
        _eState := E_DL_ElsPhase.eRamp;         (* 四站就绪 → 偏置斜坡 / All ready, ramp *)
    END_IF
E_DL_ElsPhase.eRamp:
    IF NOT xEnable THEN
        _eState := E_DL_ElsPhase.eIdle;         (* 使能撤销 → 待机 / Enable dropped *)
    ELSIF _bRampDone THEN
        _eState := E_DL_ElsPhase.eSynced;       (* 斜坡到位 → 同步相 / Ramps done, synced *)
    END_IF
E_DL_ElsPhase.eSynced:
    IF NOT xEnable THEN
        _eState := E_DL_ElsPhase.eIdle;         (* 使能撤销 → 待机 / Enable dropped *)
    ELSIF _nOnline < DL_ELS_SNUM THEN
        _eState := E_DL_ElsPhase.eEnable;       (* 从站掉线 → 回核查 / Slave offline *)
    END_IF
E_DL_ElsPhase.eFault:
    _bLimBad := FALSE;                          (* 故障相驻留：越限判据不再重算（锁存回放） *)
ELSE
    _bReqFault := TRUE;                         (* 非法相兜底 / Illegal phase fallback *)
    _eState := E_DL_ElsPhase.eFault;
END_CASE
(* 相位广播推进：仅在同步类相位推进主轴相位（eEnable/eIdle 不推进） *)
IF (_eState = E_DL_ElsPhase.eRamp) OR (_eState = E_DL_ElsPhase.eSynced) THEN
    _fMasterPhaseDeg := _fMasterPhaseDeg + _fAdvDeg;
    IF _fMasterPhaseDeg >= DL_ELS_FULL THEN
        _fMasterPhaseDeg := _fMasterPhaseDeg - DL_ELS_FULL;   (* 环绕归一 / Wrap *)
    END_IF
END_IF
(* —— 段 6：故障请求统一落地（唯一锁存点 + 同步迁相，R187/R252） —— *)
IF _bReqFault AND (NOT _bFaultLatch) THEN
    _bFaultLatch := TRUE;                       (* 锁存 / Latch *)
    _eState := E_DL_ElsPhase.eFault;            (* 同步迁相 / Migrate to fault *)
    FOR _nI := 1 TO DL_ELS_SNUM DO
        _afVelRef[_nI] := 0.0;                  (* 越限即拒并使能：速度给定全零 / All refs zero *)
    END_FOR
END_IF
(* —— 段 7：统一出口（数组在出口循环单点写入） —— *)
FOR _nI := 1 TO DL_ELS_SNUM DO
    anSlaveVelRefRpm[_nI] := _afVelRef[_nI];
END_FOR
xAllSynced := (_eState = E_DL_ElsPhase.eSynced) AND _bRampDone
              AND (_nOnline = DL_ELS_SNUM) AND (NOT _bFaultLatch) AND (NOT _bLimBad);
nSlaveOnline := _nOnline;
xFault := _bFaultLatch;
END_FUNCTION_BLOCK

(* ---- FB_DL_ExternalEncoderLatch.st ---- *)
(*==============================================================================
 * 组件名称 (Component)  : FB_DL_ExternalEncoderLatch
 * 所属子库 (Sublibrary) : DL_Motion
 * 前缀     (Prefix)     : FB_DL_
 * 当前版本 (Version)    : 1.0.0
 * 兼容性   (Platform)   : CODESYS 3.5 / TwinCAT 3 / 汇川 InoProShop / Schneider
 *                         Machine Expert；纯 IEC 61131-3（第 3 版），
 *                         仅依赖标准库 R_TRIG / F_TRIG / TON 与库内契约
 *                         I_DL_ExternalEncoder / ST_DL_EncSnapshot（只引用
 *                         不重声明），零厂商方言
 * 作者     (Author)     : 道莅代码库 · PLC编程专家（R31）
 * 开源溯源 (Origin)     : 外部编码器快照采样锁存公开语义（T1-6 外部编码器
 *                         族成员），道莅 clean-room 防御性实现，
 *                         未复制任何外部源码行
 * 功能描述 (Function)   : 外部编码器快照采样锁存件。触发上升沿调
 *                         I_DL_ExternalEncoder.Sample 写入单拍一致快照；
 *                         每拍比对当前位置与锁存位置差超容差且过期时间到
 *                         置 bStale 提示；清锁存仅由 bEn 下降沿或 bRst
 *                         复位沿显式执行，其余任何路径不得清锁存。
 *                         不自造不消费任何轴状态枚举（T1-6/MCX 家族高危区
 *                         纪律）。
 * 职责边界 (Boundary)   : 与 FB_DL_MarkPositionLatch 分工——Mark 件为轴内
 *                         探针（TouchProbe）硬件锁存，本件为外部编码器接口
 *                         的软件采样锁存，二者不合并、不互替。
 * 码位     (Codes)      : 16#0004_0067 监视级：编码器接口空引用
 *                         16#0004_0068 监视级：采样调用返回失败（保持旧值）
 *                         16#0004_0069 监视级：快照非有限拒绝入库
 *                         16#0004_006A 监视级：锁存数据过期提示（bStale）
 *                         16#0004_006B 保留未启用（码表与实现对齐，不虚声明）
 *                         本件为监视件，无 bError 出口，全码位不配故障标志。
 * 边界防错 (Boundary)   : 1 空引用判据用接口引用不等于零值判定；
 *                         2 R_TRIG/F_TRIG/TON 实例每拍无条件刷新；
 *                         3 采样失败本拍保持旧锁存值，绝不写半截快照；
 *                         4 非有限快照（x<>x 自反判加幅值界）拒绝入库；
 *                         5 bStale 为提示级，不锁存、不置故障标志。
 * 规格偏离 (Deviation)   : 规格「Reset 显式清锁存」以 bRst 复位引脚承载
 *                         （可增引脚裁定）：方法 POU 无法满足终结符纪律
 *                         中 POU 终结语句位于文件末行的要求，
 *                         引脚方案语义等价且跨平台语法风险为零。
 * 修订历史 (Revision)   : 2026-11-18 v1.0.0 首版入库（R31 · 阶段三 · 序 6）
 *==============================================================================*)

(*==============================================================================
 * 功能块: FB_DL_ExternalEncoderLatch
 * 调用约定: 每个扫描周期无条件调用一次；iEnc 引脚注入契约接口引用。
 *==============================================================================*)
FUNCTION_BLOCK FB_DL_ExternalEncoderLatch
VAR_INPUT
    iEnc      : I_DL_ExternalEncoder;       // 外部编码器契约引用（只读位置源）/ External encoder contract reference
    bTrig     : BOOL := FALSE;              // 采样触发，上升沿有效 / Sampling trigger, rising edge active
    bEn       : BOOL := FALSE;              // 使能，下降沿显式清锁存 / Enable, falling edge clears latch
    bRst      : BOOL := FALSE;              // 复位沿显式清锁存 / Reset edge clears latch explicitly
    tStale    : TIME := T#1S;               // 过期判据时长 [毫秒] / Stale judgement duration [ms]
    fPosTol   : LREAL := 0.001;             // 过期比对位置容差 [毫米] / Position tolerance for stale check [mm]
END_VAR
VAR_OUTPUT
    stLatch   : ST_DL_EncSnapshot;          // 锁存快照（同拍一致）/ Latched snapshot, scan-consistent
    bLatchValid : BOOL;                     // 锁存有效标志 / Latch validity flag
    bStale    : BOOL;                       // 锁存数据过期提示 / Stale data notice
    uErrorId  : UDINT;                      // 监视级码，0 = 无（段位码需 32 位载体）/ Monitor code, 0 = none, segment codes need 32-bit
END_VAR
VAR
    rTrigTrig : R_TRIG;                     // 采样触发沿检测，每拍无条件刷新 / Trigger edge detector, refreshed every scan
    fTrigEn   : F_TRIG;                     // 使能下降沿检测，每拍无条件刷新 / Enable falling edge detector
    rTrigRst  : R_TRIG;                     // 复位沿检测，每拍无条件刷新 / Reset edge detector, refreshed every scan
    tonStale  : TON;                        // 过期计时器，每拍无条件刷新 / Stale timer, refreshed every scan
    stTmp     : ST_DL_EncSnapshot;          // 采样暂存快照 / Sampling temp snapshot
    fNowPos   : LREAL;                      // 本拍当前位置 [毫米] / Current position this scan [mm]
    bEncOk    : BOOL;                       // 接口引用有效标志 / Interface reference valid flag
    bSampleOk : BOOL;                       // 本拍采样受理标志 / Sampling accepted flag this scan
    bSnapOk   : BOOL;                       // 快照有限有效标志 / Snapshot finiteness flag
    xRstOne   : BOOL;                       // 过期计时单拍重置请求 / One-scan stale timer reset request
END_VAR
VAR CONSTANT
    DL_EEL_FIN : LREAL := 1.0E30;           // LREAL 有限幅值判界 / LREAL finiteness magnitude bound
END_VAR

// ---- 段 1｜边沿与定时器实例无条件周期刷新（红线：禁入条件分支）----------------
rTrigTrig(CLK := bTrig);                                 // 触发沿检测 / Trigger edge detection
fTrigEn(CLK := bEn);                                     // 使能下降沿检测 / Enable falling edge detection
rTrigRst(CLK := bRst);                                   // 复位沿检测 / Reset edge detection
tonStale(IN := (bLatchValid AND bEn AND NOT xRstOne), PT := tStale); // 过期计时 / Stale timing

// ---- 段 2｜接口引用有效性与当前位置读取 ----------------------------------------
bEncOk := (iEnc <> 0);                                   // 接口引用非空判定 / Interface reference not null
IF bEncOk THEN
    fNowPos := iEnc.fPos;                                // 读当前位置 [毫米] / Read current position
ELSE
    fNowPos := 0.0;                                      // 空引用确定值 / Deterministic fallback
END_IF

// ---- 段 3｜清锁存唯一通道：使能下降沿、复位沿（两路显式，别无路径）--------------
IF fTrigEn.Q OR rTrigRst.Q THEN
    bLatchValid := FALSE;                                // 显式清锁存 / Explicit latch clear
    stLatch.fPos := 0.0;                                 // 快照位置清零 / Zero snapshot position
    stLatch.fVel := 0.0;                                 // 快照速度清零 / Zero snapshot velocity
    stLatch.tStamp := T#0MS;                             // 快照时戳清零 / Zero snapshot timestamp
    stLatch.bValid := FALSE;                             // 快照有效位清零 / Zero snapshot validity
    bStale := FALSE;                                     // 清过期提示 / Clear stale notice
END_IF

// ---- 段 4｜触发沿采样入库 -------------------------------------------------------
bSampleOk := FALSE;                                      // 受理标志先清 / Clear accepted flag
bSnapOk := FALSE;                                        // 有限标志先清 / Clear finiteness flag
IF bEncOk AND bEn AND rTrigTrig.Q THEN
    bSampleOk := iEnc.Sample(stSnap := stTmp);           // 调契约采样方法 / Invoke contract sampling method
    IF bSampleOk THEN
        bSnapOk := (stTmp.fPos = stTmp.fPos) AND (stTmp.fVel = stTmp.fVel)
               AND (ABS(stTmp.fPos) < DL_EEL_FIN) AND (ABS(stTmp.fVel) < DL_EEL_FIN); // 快照双字段有限 / Both fields finite
        IF bSnapOk THEN
            stLatch     := stTmp;                        // 快照整体入库 / Snapshot committed
            bLatchValid := TRUE;                         // 锁存有效 / Latch valid
            xRstOne     := TRUE;                         // 单拍断过期计时输入 / One-scan stale timer break
        END_IF                                           // 非有限拒绝入库保持旧值 / Non-finite rejected, keep old
    END_IF                                               // 采样失败保持旧锁存 / Sampling failed, keep old latch
END_IF

// ---- 段 5｜过期提示判定：过期时长到且位置差超容差 -------------------------------
bStale := tonStale.Q AND bLatchValid
      AND (ABS(fNowPos - stLatch.fPos) > fPosTol);       // 过期与漂移双条件 / Stale duration and drift both required

// ---- 段 6｜监视级码装配（监视件不置故障标志）------------------------------------
IF NOT bEncOk THEN
    uErrorId := 16#0004_0067;                            // 空引用码 / Null reference code
ELSIF bEncOk AND bEn AND rTrigTrig.Q AND (NOT bSampleOk) THEN
    uErrorId := 16#0004_0068;                            // 采样失败码 / Sampling failure code
ELSIF bEncOk AND bEn AND rTrigTrig.Q AND bSampleOk AND (NOT bSnapOk) THEN
    uErrorId := 16#0004_0069;                            // 快照非有限码 / Non-finite snapshot code
ELSIF bStale THEN
    uErrorId := 16#0004_006A;                            // 过期提示码 / Stale notice code
ELSE
    uErrorId := 16#0000_0000;                            // 无码 / No code
END_IF

// ---- 段 7｜单拍标志收尾 ----------------------------------------------------------
xRstOne := FALSE;                                        // 重置请求仅当拍有效 / Reset request is single scan
END_FUNCTION_BLOCK

(* ---- FB_DL_ExternalEncoderScaler.st ---- *)
(*
    FB_DL_ExternalEncoderScaler —— 外部编码器折算
    ------------------------------------------------------------------
    分类      : DL_Motion / Feedback
    前缀      : FB_DL_
    版本      : 1.0.0
    溯源      : 只借「外部编码器属运动层反馈、可独立成块」的分类事实（公开运动控制示例
                的组织划分）；回绕展开算法、折算链顺序、错误分级与码位 100% 自有；
                本件不自造轴状态、不发运动指令、不消费任何厂商轴接口；
                clean-room 重写，未复制任何闭源厂商源码
    平台      : 纯 IEC 61131-3，CODESYS V3.5+ / TwinCAT 3 / InoProShop 通用
    作者      : 道莅代码库 · PLC编程专家（R19）
    ------------------------------------------------------------------
    功能说明  : 把外部编码器原始计数折算成工程量（mm / 度），含分辨率、传动比、导程三段
                折算与 32 位计数器回绕展开（不展开则多圈坐标每转一圈就跳变）。
                **本件最易错的一行**：回绕判据必须先做 DINT 减法、再升位到 LINT——
                先升位再减会让 32 位回绕变成巨大正数（R68 硬纪律）。
                其余防御：① 分辨率或导程为 0 即故障级（除零唯一出口），输出冻结；
                ② 传动比分子或分母为 0 即故障级 02DF；
                ③ 计数器位宽越域只钳位并置信息码（钳位后回绕判据仍可用，不必停功能）；
                ④ 首拍只装初值、不产生回绕事件；
                ⑤ 折算结果非有限即故障级并保持末次有效位置——掉成 0 会被上层当成真实回零。
                规格补正：fVelocity [mm/s] 需要时间基准，派单未给采样周期引脚，特补
                tSampleTime（否则速度只能伪造），收口报告留档。
                职责边界：卷径/张力等工艺量归各自工艺件，本件只出位置与速度。
    错误码    : 16#0004_01CD 检测到计数回绕已展开 / 位宽参数超域已钳位——信息级，正常防御
                16#0004_01CE 预留禁用（信息级，不得挪用）
                16#0004_02DE 分辨率或导程非法（为 0 / 非有限）——故障级，输出冻结
                16#0004_02DF 传动比分子或分母为 0——故障级，输出冻结
                16#0004_02E0 折算结果非有限——故障级，保持末次有效位置
    码位总账  : 16#0004_01CD 用 / 16#0004_01CE 预留 ｜ 16#0004_02DE 用 / 16#0004_02DF 用 / 16#0004_02E0 用
    状态机    : R6 标注 N/A —— 本组件为纯函数无顺序状态机，无 CASE 可写，非法状态不可能出现
                （首拍由单比特 bInit 承载，非顺序状态机）
    采样约定  : fbTrigReset 在本体首部无条件刷新；速度由相邻拍位置差分除以 tSampleTime 得到，
                采样周期为 0 时速度置 0（不做除零），位置折算与之无关。
    修订记录  : 2026-11-16 v1.0.0 首次入库（R19）
*)
FUNCTION_BLOCK FB_DL_ExternalEncoderScaler
VAR_INPUT
    bEnable         : BOOL;                   // 使能，FALSE 输出冻结 / enable, FALSE freezes the outputs
    bReset          : BOOL;                   // 复位，上升沿清多圈展开与零点 / reset, rising edge clears the multi-turn unfolding and the datum
    diRawCount      : DINT := 0;              // 原始计数（编码器直接读出的 32 位值）[count] / raw count read from the encoder [count]
    uCountsPerRev   : UDINT := 4096;          // 每转计数 [count/rev]，必须 > 0 / counts per revolution [count/rev], must be > 0
    fPitch          : REAL := 5.0;            // 每转行程（丝杠导程 / 辊周长）[mm/rev]，必须 > 0 / travel per revolution [mm/rev], must be > 0
    iGearNum        : INT := 1;               // 传动比分子 [无量纲]，必须 != 0 / gear ratio numerator [dimensionless], must be nonzero
    iGearDen        : INT := 1;               // 传动比分母 [无量纲]，必须 != 0 / gear ratio denominator [dimensionless], must be nonzero
    bInvert         : BOOL := FALSE;          // TRUE = 方向取反 / TRUE inverts the direction
    fOffset         : REAL := 0.0;            // 零点偏置 [mm] / datum offset [mm]
    nMultiTurnBits  : INT := 32;              // 计数器位宽 [bit]，范围 8~32 / counter width [bit], range 8~32
    tSampleTime     : TIME := T#10MS;         // 采样周期（规格补正引脚，速度折算用）[ms]，范围 1~1000 / sample time, a spec correction pin used by the velocity conversion [ms], range 1~1000
END_VAR
VAR_OUTPUT
    fPosition       : REAL;                   // 折算后工程量 [mm] / converted engineering position [mm]
    liTotalCount    : LINT;                   // 展开后的多圈累计计数 [count] / unfolded multi-turn accumulated count [count]
    bWrapped        : BOOL;                   // 本拍检测到回绕（单周期脉冲）/ a wrap was detected in this cycle, single-cycle pulse
    uWrapCount      : UDINT;                  // 累计回绕次数，饱和 [次] / accumulated wrap count, saturating [times]
    fVelocity       : REAL;                   // 相邻拍差分估计速度（仅供监视）[mm/s] / velocity estimated from consecutive cycles, monitoring only [mm/s]
    eErr            : UDINT;                  // 错误码，0=正常 / error id, 0=ok
    bError          : BOOL;                   // 故障标志，eErr 为故障级时 TRUE / error flag, TRUE on fault-level eErr
    bValid          : BOOL;                   // 输出是否可用 / output valid flag
END_VAR
VAR
    fbTrigReset     : R_TRIG;                 // 复位上升沿实例，本体首部无条件刷新 / reset edge instance, refreshed unconditionally
    diPrevRaw       : DINT;                   // 上一拍原始计数 [count] / previous raw count [count]
    liAccum         : LINT;                   // 多圈累计计数 [count] / multi-turn accumulated count [count]
    liDelta         : LINT;                   // 单拍计数增量（升位后）[count] / per cycle increment widened to LINT [count]
    liHalfSpan      : LINT;                   // 半量程（2^(位宽-1)）[count] / half span of the counter [count]
    liFullSpan      : LINT;                   // 全量程（2^位宽）[count] / full span of the counter [count]
    nDelta          : DINT;                   // 单拍计数增量（先做 DINT 减法）[count] / per cycle increment computed in DINT first [count]
    nBitsEff        : INT;                    // 钳位后的计数器位宽 [bit] / clamped counter width [bit]
    fRatio          : REAL;                   // 圈数（含小数）[rev] / revolution count including the fraction [rev]
    fGear           : REAL;                   // 传动比（分子/分母）[无量纲] / gear ratio, numerator over denominator [dimensionless]
    fSign           : REAL;                   // 方向符号 [+1 / -1] / direction sign, plus or minus one
    fPos            : REAL;                   // 折算位置中间量 [mm] / converted position intermediate [mm]
    fDtSec          : REAL;                   // 采样周期秒值 [s] / sample time in seconds [s]
    fPrevPos        : REAL;                   // 上一拍位置 [mm] / previous position [mm]
    bInit           : BOOL := FALSE;          // 首扫标志，初值 FALSE，判据 NOT bInit / first-scan flag, initial FALSE, tested with NOT
    nDtMs           : DINT;                   // 采样周期毫秒整数 [ms] / sample time in integer milliseconds [ms]
END_VAR
VAR CONSTANT
    DL_EES_CPR_MIN   : UDINT := 1;            // 每转计数下限 [count/rev] / counts per revolution lower bound [count/rev]
    DL_EES_BITS_MIN  : INT := 8;              // 计数器位宽下限 [bit] / counter width lower bound [bit]
    DL_EES_BITS_MAX  : INT := 32;             // 计数器位宽上限 [bit] / counter width upper bound [bit]
    DL_EES_CNT_MAX   : UDINT := 16#FFFF_FFFE; // 回绕计数饱和值 [次] / wrap counter saturation value [times]
    DL_EES_DT_MIN    : TIME := T#1MS;         // 采样周期下限 [ms] / sample time lower bound [ms]
    DL_EES_DT_MAX    : TIME := T#1S;          // 采样周期上限 [ms] / sample time upper bound [ms]
    DL_FLOAT_EPS     : REAL := 1.0E-6;        // 浮点判等容差 [无量纲] / float equality tolerance [dimensionless]
    DL_EES_INF_GUARD : REAL := 1.0E38;        // 非有限幅值判定阈值 [无量纲] / non-finite magnitude guard [dimensionless]
    DL_EES_MS_PER_S  : REAL := 1000.0;        // 毫秒到秒换算因子 [ms/s] / milliseconds per second [ms/s]
    DL_EES_TWO       : LINT := 2;             // 整型二值常量，量程倍数用 [无量纲] / integer two used for the span multiples
    DL_EES_ONE       : LINT := 1;             // 整型一值常量，位运算基底 [无量纲] / integer one used as the shift base
    DL_EES_SIGN_POS  : REAL := 1.0;           // 正向符号 [+1] / positive direction sign
    DL_EES_SIGN_NEG  : REAL := -1.0;          // 反向符号 [-1] / negative direction sign
    DL_EES_ZERO      : REAL := 0.0;           // 零值常量，避免裸字面量 [无量纲] / zero constant, avoids a bare literal [dimensionless]
    DL_EES_ZERO_L    : LINT := 0;             // LINT 零值常量 [count] / LINT zero constant [count]
    DL_EES_ZERO_U    : UDINT := 0;            // UDINT 零值常量 [无量纲] / UDINT zero constant [dimensionless]
END_VAR

// 段 1｜边沿实例无条件周期刷新（红线：严禁放入条件分支）/ segment 1, unconditional edge refresh
fbTrigReset(CLK := bReset);

// 段 2｜输出与错误状态预置（fPosition / liTotalCount 为保持量，故障时须保末值）/ segment 2, preset outputs, the held values are kept
eErr := 0;                                    // 预置无错误 / preset no error
bError := FALSE;                              // 预置无故障 / preset no fault
bValid := FALSE;                              // 预置不可用 / preset invalid
bWrapped := FALSE;                            // 单周期脉冲先清 / clear the single-cycle pulse

// 段 3｜参数闸一：分辨率与导程（除零唯一出口）/ segment 3, resolution and pitch gate
IF (uCountsPerRev < DL_EES_CPR_MIN)
   OR (fPitch <= DL_FLOAT_EPS)
   OR (fPitch <> fPitch) OR (fPitch > DL_EES_INF_GUARD) OR (fPitch < -DL_EES_INF_GUARD) THEN
    eErr := 16#0004_02DE;                     // 分辨率或导程非法故障码 / resolution or pitch fault id
    bError := TRUE;                           // 置故障标志 / raise the error flag
    bValid := FALSE;                          // 输出冻结 / the output stays frozen
    RETURN;                                   // 故障级提前返回，不进入任何除法 / early return before any division
END_IF

// 段 4｜参数闸二：传动比分子分母非零 / segment 4, gear ratio gate
IF (iGearNum = 0) OR (iGearDen = 0) THEN
    eErr := 16#0004_02DF;                     // 传动比为 0 故障码 / zero gear ratio fault id
    bError := TRUE;                           // 置故障标志 / raise the error flag
    bValid := FALSE;                          // 输出冻结 / the output stays frozen
    RETURN;                                   // 故障级提前返回 / early return on fault
END_IF

// 段 5｜位宽钳位（钳位后回绕判据仍可用，不必停功能）/ segment 5, width clamping
nBitsEff := nMultiTurnBits;                   // 取入参副本 / copy the input
IF nBitsEff < DL_EES_BITS_MIN THEN
    nBitsEff := DL_EES_BITS_MIN;              // 位宽下限钳位 / clamp at the lower bound
    eErr := 16#0004_01CD;                     // 信息级：位宽超域已钳位 / info level, the width was clamped
ELSIF nBitsEff > DL_EES_BITS_MAX THEN
    nBitsEff := DL_EES_BITS_MAX;              // 位宽上限钳位 / clamp at the upper bound
    eErr := 16#0004_01CD;                     // 信息级：位宽超域已钳位 / info level, the width was clamped
END_IF

// 段 6｜半量程与全量程（LINT 承载，避开 2^31 在 DINT 域溢出）/ segment 6, half and full span in LINT
liHalfSpan := SHL(DL_EES_ONE, nBitsEff - 1);  // 2^(位宽-1)，移位量 <= 31 结构性安全 / two to the width minus one, the shift never exceeds 31
liFullSpan := liHalfSpan * DL_EES_TWO;        // 2^位宽 / two to the width

// 段 7｜使能闸：失能冻结输出 / segment 7, enable gate freezes the outputs
IF NOT bEnable THEN
    RETURN;                                   // 失能即出口，输出保持 / disabled is the exit, the outputs are held
END_IF

// 段 8｜首扫初始化：只装初值，不产生回绕事件 / segment 8, first-scan initialisation without a wrap event
IF NOT bInit THEN
    liAccum := DL_EES_ZERO_L;                 // 累计计数清零 / clear the accumulated count
    diPrevRaw := diRawCount;                  // 原始计数基准装载 / load the raw count reference
    fPrevPos := fOffset;                      // 位置基准取偏置 / the position reference starts at the offset
    uWrapCount := DL_EES_ZERO_U;              // 回绕计数清零 / clear the wrap counter
    bInit := TRUE;                            // 首扫只做一次 / first scan runs once only
    fPosition := fOffset;                     // 首拍位置即偏置 / the first position equals the offset
    liTotalCount := liAccum;                  // 首拍累计计数输出 / publish the accumulated count
    bValid := TRUE;                           // 首拍输出可用 / the first scan output is usable
    RETURN;                                   // 首拍不做回绕判定 / no wrap detection on the first scan
END_IF

// 段 9｜复位沿：清多圈展开与零点基准 / segment 9, reset clears the unfolding and the datum
IF fbTrigReset.Q THEN
    liAccum := DL_EES_ZERO_L;                 // 累计计数清零 / clear the accumulated count
    diPrevRaw := diRawCount;                  // 基准重装 / reload the reference
    fPrevPos := fOffset;                      // 位置基准回偏置 / the position reference returns to the offset
    uWrapCount := DL_EES_ZERO_U;              // 回绕计数清零 / clear the wrap counter
END_IF

// 段 10｜回绕展开（R68 硬纪律：先做 DINT 减法，再升位比较）/ segment 10, wrap unfolding, subtract first then widen
nDelta := diRawCount - diPrevRaw;             // 先做 32 位减法：回绕在此自然发生 / the 32-bit subtraction comes first, the wrap happens here naturally
diPrevRaw := diRawCount;                      // 立即更新基准 / update the reference immediately
liDelta := DINT_TO_LINT(nDelta);              // 减法之后才升位，顺序不可颠倒 / widen only after the subtraction
IF liDelta > liHalfSpan THEN
    liDelta := liDelta - liFullSpan;          // 正向回绕展开 / unfold a forward wrap
    bWrapped := TRUE;                         // 标记回绕事件 / flag the wrap event
ELSIF liDelta < -liHalfSpan THEN
    liDelta := liDelta + liFullSpan;          // 反向回绕展开 / unfold a backward wrap
    bWrapped := TRUE;                         // 标记回绕事件 / flag the wrap event
END_IF
liAccum := liAccum + liDelta;                 // 累计计数（LINT 域，长期不溢出）/ accumulate in the LINT domain, no overflow in practice

// 段 11｜回绕计数与信息码 / segment 11, wrap counter and info code
IF bWrapped THEN
    IF uWrapCount < DL_EES_CNT_MAX THEN
        uWrapCount := uWrapCount + 1;         // 饱和加一 / saturating increment
    END_IF
    eErr := 16#0004_01CD;                     // 信息级：检测到回绕已展开 / info level, a wrap was detected and unfolded
END_IF

// 段 12｜三段折算链（分母已由段 3 / 段 4 保证非零）/ segment 12, three stage conversion chain
fRatio := LINT_TO_REAL(liAccum) / UDINT_TO_REAL(uCountsPerRev); // 圈数（含小数）[rev] / revolutions including the fraction [rev]
fGear := INT_TO_REAL(iGearNum) / INT_TO_REAL(iGearDen);         // 传动比 [无量纲] / gear ratio [dimensionless]
IF bInvert THEN
    fSign := DL_EES_SIGN_NEG;                 // 方向取反 / invert the direction
ELSE
    fSign := DL_EES_SIGN_POS;                 // 方向保持 / keep the direction
END_IF
fPos := fRatio * fPitch * fGear * fSign + fOffset; // 位置折算 [mm] / convert to the engineering position [mm]

// 段 13｜结果非有限闸：保持末次有效位置（掉成 0 会被当成真实回零）/ segment 13, non-finite gate holds the last position
IF (fPos <> fPos) OR (fPos > DL_EES_INF_GUARD) OR (fPos < -DL_EES_INF_GUARD) THEN
    eErr := 16#0004_02E0;                     // 折算结果非有限故障码 / non-finite conversion fault id
    bError := TRUE;                           // 置故障标志 / raise the error flag
    bValid := FALSE;                          // 输出不可用 / the output is not usable
    RETURN;                                   // fPosition 保持末次有效值 / fPosition keeps its last valid value
END_IF

// 段 14｜速度差分（采样周期为 0 时置 0，不做除零）/ segment 14, velocity by difference with a guarded divisor
nDtMs := TIME_TO_DINT(tSampleTime);           // 采样周期整数毫秒 [ms] / sample time in integer milliseconds [ms]
IF (nDtMs > 0) AND (tSampleTime >= DL_EES_DT_MIN) AND (tSampleTime <= DL_EES_DT_MAX) THEN
    fDtSec := DINT_TO_REAL(nDtMs) / DL_EES_MS_PER_S; // 换算为秒 [s] / convert to seconds [s]
    fVelocity := (fPos - fPrevPos) / fDtSec;  // 差分速度 [mm/s] / differential velocity [mm/s]
ELSE
    fVelocity := DL_EES_ZERO;                 // 周期非法则速度不可信，输出 0 / an illegal period makes the velocity untrustworthy, output zero
END_IF

// 段 15｜发布结果 / segment 15, publish the results
fPosition := fPos;                            // 输出折算位置 [mm] / publish the converted position [mm]
liTotalCount := liAccum;                      // 输出多圈累计计数 [count] / publish the accumulated count [count]
fPrevPos := fPos;                             // 记录为下一拍差分基准 / remember it for the next difference
bValid := TRUE;                               // 通过全部闸门，输出可用 / all gates passed, the output is usable
bError := FALSE;                              // 信息级不置故障 / info level never raises a fault
END_FUNCTION_BLOCK

(* ---- FB_DL_FeedOverrideRamp.st ---- *)
(*
  ==================================================================
  组件名 Component  : FB_DL_FeedOverrideRamp
  分类   Category   : DL_Motion
  前缀   Naming     : FB_DL_ ｜ b/n/u/f/t/e 类型前缀制（R265）
  版本   Version    : 1.0.0
  功能   Purpose    : 进给倍率斜坡（PLCopen 风格 0~150%）：正常相按「加速/
                      减速」分离速率把 fOvrOut 斜坡逼近钳位后的 fOvrIn；
                      bZeroFast 为显式最高优先级仲裁——TRUE 时无条件以
                      fRateZeroPctS 向 0% 斜坡（压倒正常跟踪）；bAtCmd 用
                      1E-6 容差判到达（禁浮点判等）。
  来源   Source     : t1-6-plcopen（PLCopen TC 系列倍率语义：借「倍率域与
                      速率限制」公开口径，实现零源码复制）
  互引   Cross-ref  : FB_DL_RateLimiter（同族通用限速率器，本件为其倍率域
                      特化件，速率仲裁口径一致）；FB_DL_OverrideSelector
                      （上游倍率源选择件，其输出可接本件 fOvrIn）
  平台   Platform   : 纯 IEC 61131-3 四则，三平台通用
  依赖   Depends    : 无标准库依赖（无定时器/无沿检测）
  设计偏差 Deviation: 时间基准按本库「时间注入」纪律：新增输入 fCallCycleS
                      （调用方注入扫描周期 [s]），本件不读平台时刻函数；
                      斜坡步长 = 速率 × fCallCycleS。
  红线   Redline    : R1 零全局/VAR_EXTERNAL/R2 零 %I/%Q/R3 纯 IEC 标准
                      R4 输入 0~150 显式钳位 + 输出 0~150 显式钳位 +
                      非有限闸 + 容差判到达（禁 =）+ 除法零处（无除法面）
                      R5 全变量双语同行注释/R6 纯仲裁无 ENUM 状态机（仲裁
                      优先级线性结构，非相态迁移，见头注说明）
                      R7 无定时器与沿检测实例/R8 速率与容差常量化
  契约   Contract   : 失能相输出行为写死（FB33-4 声明，不静默）：bEnable=
                      FALSE → fOvrOut 冻结保持上次值、bAtCmd=FALSE，速率
                      配置不复检（恢复使能后重新生效）；bZeroFast 使能独立
                      于 bEnable（安全归零不受失能门控压制，头注安全侧口径）。
  错误码 Codes      : 01【故障级】速率配置非法（fRateIncPctS / fRateDecPctS /
                      fRateZeroPctS 任一 ≤ 0 或非有限，或 fCallCycleS ≤ 0 /
                      非有限）；故障相输出冻结保持 + bError（R45 配对）
  码位反证 Note     : 仅一码依据（R90 反证）：三个速率任一非法的处置完全
                      同形（冻结 + 拒斜坡），输出组合不可区分，合并不丢信息。
  验收   Acceptance : V1 30→80% 增速斜坡按 fRateIncPctS ｜ V2 80→30% 按
                      fRateDecPctS ｜ V3 bZeroFast → 以 fRateZeroPctS 归零，
                      bEnable=FALSE 时仍归零（仲裁显式）｜ V4 速率 0 → 码 01
                      + 冻结 ｜ V5 到达 ±1E-6 内 bAtCmd=TRUE ｜ V6 全程不出
                      [0,150]
  变更   Revision   : 2026-11-22  v1.0.0  R66 首版（编码阶段批 3 序 8）
  ==================================================================
*)
FUNCTION_BLOCK FB_DL_FeedOverrideRamp
VAR_INPUT
    fOvrIn       : LREAL := 0.0;    // 倍率请求 [%]，0~150 钳位 / the override request, clamped 0 to 150
    bEnable      : BOOL := FALSE;   // 使能（失能=冻结保持，头注契约写死）[-] / the enable, false freezes the output
    bZeroFast    : BOOL := FALSE;   // 快速归零仲裁（最高优先级，独立于使能）[-] / the fast zero arbitration, the top priority
    fRateIncPctS : LREAL := 50.0;   // 增速率 [%/s]，须 > 0 / the increase rate, must be positive
    fRateDecPctS : LREAL := 50.0;   // 减速率 [%/s]，须 > 0 / the decrease rate, must be positive
    fRateZeroPctS: LREAL := 200.0;  // 归零速率 [%/s]，须 > 0（仲裁用）/ the zero rate, must be positive
    fCallCycleS  : LREAL := 0.01;   // 调用方注入扫描周期 [s]，须 > 0 / the caller injected scan cycle in seconds
END_VAR
VAR_OUTPUT
    fOvrOut      : LREAL := 0.0;    // 倍率输出 [%]，全程钳位 0~150 / the override output, always clamped 0 to 150
    bAtCmd       : BOOL := FALSE;   // 到达指示（1E-6 容差判到达）[-] / the at command flag by tolerance
    bError       : BOOL := FALSE;   // 配置故障标志（R45 配对）/ the configuration fault flag
    uErrorId     : UDINT := 16#0000_0000; // 错误码，0=正常，01=速率配置非法 [码] / the error code [code]
END_VAR
VAR
    _fTarget     : LREAL := 0.0;    // 本拍斜坡目标 [%] / the per scan ramp target
    _fRate       : LREAL := 0.0;    // 本拍选用速率 [%/s] / the per scan selected rate
    _fStep       : LREAL := 0.0;    // 本拍斜坡步长 [%] / the per scan ramp step
    _bCfgOk      : BOOL := FALSE;   // 本拍配置有效性 [-] / the per scan configuration validity
END_VAR
VAR CONSTANT
    FOR_OVR_MIN  : LREAL := 0.0;      // 倍率域下限 [%] / the override domain lower clamp
    FOR_OVR_MAX  : LREAL := 150.0;    // 倍率域上限 [%]（PLCopen 倍率域口径）/ the override domain upper clamp
    FOR_AT_EPS   : LREAL := 1.0E-6;   // 到达容差 [%]（禁浮点判等）/ the arrival tolerance
    FOR_FIN_MAX  : LREAL := 1.7976931348623157E308; // LREAL 有限上限 / the finite LREAL limit
    FOR_ERR_NONE : UDINT := 16#0000_0000; // 无错误 [码] / no error [code]
    FOR_ERR_RATE : UDINT := 16#0000_0001; // 码 01：速率配置非法 / code 01, illegal rate configuration
END_VAR

// 段 1｜配置闸（码 01）：三速率与扫描周期逐项有限 + 正域 / segment 1, the configuration gate
_bCfgOk := (fRateIncPctS > 0.0) AND (fRateIncPctS = fRateIncPctS)
       AND (fRateDecPctS > 0.0) AND (fRateDecPctS = fRateDecPctS)
       AND (fRateZeroPctS > 0.0) AND (fRateZeroPctS = fRateZeroPctS)
       AND (fCallCycleS > 0.0) AND (fCallCycleS = fCallCycleS);   // 逐项自反判 NaN + 正域 / per item NaN reflex and positivity
IF _bCfgOk THEN
    bError := FALSE;                 // 配置恢复即清标志（信息级随当拍，无锁存面）/ cleared when the config recovers
    uErrorId := FOR_ERR_NONE;
ELSE
    bError := TRUE;                  // 故障标志（R45 配对）/ the fault flag
    uErrorId := FOR_ERR_RATE;        // 码 01 / code 01
    bAtCmd := FALSE;                 // 故障相到达指示撤销（头注契约）/ revoke the arrival flag in the fault phase
    RETURN;                          // 故障相输出冻结保持 fOvrOut（头注契约），不再斜坡 / frozen output, no ramping
END_IF

// 段 2｜请求钳位与非有限闸：非有限请求按 0% 安全侧处理 / segment 2, the request clamp and finiteness gate
IF (fOvrIn <> fOvrIn) OR (ABS(fOvrIn) > FOR_FIN_MAX) THEN
    _fTarget := FOR_OVR_MIN;         // 非有限请求落 0%（安全侧）/ a non finite request lands at zero
ELSIF fOvrIn < FOR_OVR_MIN THEN
    _fTarget := FOR_OVR_MIN;         // 下钳 / clamp low
ELSIF fOvrIn > FOR_OVR_MAX THEN
    _fTarget := FOR_OVR_MAX;         // 上钳 / clamp high
ELSE
    _fTarget := fOvrIn;              // 合法请求直取 / take the valid request
END_IF

// 段 3｜归零优先仲裁（显式优先序：bZeroFast > bEnable 跟踪，线性仲裁无状态相）
//      segment 3, the explicit arbitration, zero fast outranks the tracking
IF bZeroFast THEN
    _fTarget := FOR_OVR_MIN;         // 归零目标（压倒请求）/ the zero target overrides the request
    _fRate := fRateZeroPctS;         // 归零专用速率 / the dedicated zero rate
ELSIF NOT bEnable THEN
    bAtCmd := FALSE;                 // 失能相到达指示撤销（头注契约写死）/ revoke the arrival flag in the disabled phase
    RETURN;                          // 失能相：输出冻结保持 fOvrOut（头注契约写死）/ the disabled phase freezes
ELSE
    IF fOvrOut < _fTarget THEN
        _fRate := fRateIncPctS;      // 向上用增速率 / the increase rate upward
    ELSE
        _fRate := fRateDecPctS;      // 向下用减速率 / the decrease rate downward
    END_IF
END_IF

// 段 4｜斜坡推进（步长 = 速率 × 周期，周期已闸 > 0）/ segment 4, the ramp advance
_fStep := _fRate * fCallCycleS;      // 本拍步长 [%] / the per scan step
IF fOvrOut < _fTarget - FOR_AT_EPS THEN
    fOvrOut := fOvrOut + _fStep;     // 向上斜坡 / ramp up
    IF fOvrOut > _fTarget THEN fOvrOut := _fTarget; END_IF   // 不越过目标 / never past the target
ELSIF fOvrOut > _fTarget + FOR_AT_EPS THEN
    fOvrOut := fOvrOut - _fStep;     // 向下斜坡 / ramp down
    IF fOvrOut < _fTarget THEN fOvrOut := _fTarget; END_IF
END_IF

// 段 5｜输出钳位（双保险）与到达判定 / segment 5, the output clamp and the arrival test
IF fOvrOut < FOR_OVR_MIN THEN
    fOvrOut := FOR_OVR_MIN;          // 下限钳位 / clamp low
END_IF
IF fOvrOut > FOR_OVR_MAX THEN
    fOvrOut := FOR_OVR_MAX;          // 上限钳位 / clamp high
END_IF
bAtCmd := ABS(fOvrOut - _fTarget) < FOR_AT_EPS;  // 容差判到达（禁 =）/ arrival by tolerance
END_FUNCTION_BLOCK

(* ---- FB_DL_FilmSpliceTensionHold.st ---- *)
// =====================================================================
// FB_DL_FilmSpliceTensionHold.st
// 接膜瞬间张力双回路无扰交接（给定斜坡 + 权重交叉淡入淡出）
// Film splice tension handover FB
// 码位: 16#0004_0345 ~ 16#0004_0349 (本件独占 5 槽)
// 修改记录: R29 初版 (按 DISPATCH_R29 序 13)
// =====================================================================
FUNCTION_BLOCK FB_DL_FilmSpliceTensionHold
VAR_INPUT
    bEnable       : BOOL  := FALSE;    // 使能 / Enable
    bSpliceStart  : BOOL  := FALSE;    // 上升沿启动交接 / Splice start on edge
    bReset        : BOOL  := FALSE;    // 复位 / Reset
    fTensionA_N   : REAL  := 0.0;      // A 卷实测张力 0~2000 N / A tension [N]
    fTensionANow_N: REAL  := 0.0;      // A 卷当前指令值 0~2000 N / A command [N]
    fTensionBSp_N : REAL  := 200.0;    // B 卷目标张力 0~2000 N / B setpoint [N]
    bBMeasValid   : BOOL  := FALSE;    // B 卷张力实测有效 / B measurement valid
    fRamp_Ns      : REAL  := 200.0;    // 给定斜坡速率 1~5000 N/s / Ramp rate [N/s]
    fDevMax_N     : REAL  := 40.0;     // 交接允许偏差 1~500 N / Max deviation [N]
    tHoldMax      : TIME  := T#3S;     // 交接最长时间 T#100MS~T#30S / Max handover time [s]
    tCycle        : TIME  := T#10MS;   // 周期 T#1MS~T#200MS / Cycle [s]
END_VAR
VAR_OUTPUT
    fTensionCmd_N : REAL;              // 交接后张力给定 0~2000 N / Tension command [N]
    fBlendPct     : REAL;              // B 回路权重 0~100 % / Blend weight [%]
    bHoldActive   : BOOL;              // 交接进行中 / Handover active
    bHandoverDone : BOOL;              // 交接完成（单拍脉冲）/ Handover done pulse
    bCutPermit    : BOOL;              // 允许裁切 / Cut permit
    eErr          : UDINT;             // 错误码 / Error code
END_VAR
VAR
    rtrigStart    : R_TRIG;            // 启动沿检测（无条件刷新）/ Start edge detector
    fStepN        : REAL;              // 单拍给定增量 / Step per cycle [N]
    tHoldMaxS     : REAL;              // 上限秒值 / Hold max seconds [s]
    tCycleS       : REAL;              // 周期秒值 / Cycle seconds [s]
    bHoldLatch    : BOOL := FALSE;     // 交接超时中止锁存 / Handover abort latch
    bDevFrozen    : BOOL := FALSE;     // 偏差超限冻结标志 / Deviation freeze flag
    fStartCmd     : REAL;              // 交接起始给定快照 / Handover start command snapshot [N]
    tonHold       : TON;               // 交接超时定时器（无条件刷新）/ Handover timeout timer
    xFirstScan    : BOOL  := TRUE;     // 首扫标记 / First-scan flag
END_VAR

// ---------------------------------------------------------------------
// 代码位表（本件独占，勿复用）:
//   16#0004_0345 信息 交接完成 / 未启动
//   16#0004_0346 故障 张力非有限 / tCycle 非法
//   16#0004_0347 故障 fRamp_Ns ≤ 0 / fTensionBSp_N ≤ 0 / tHoldMax 非法（组态错）
//   16#0004_0348 信息 交接中偏差超 fDevMax_N → 冻结斜坡与权重，bHoldActive 保持
//   16#0004_0349 故障 交接超 tHoldMax 未达 100 % → 中止、bCutPermit=FALSE 锁存
// ---------------------------------------------------------------------

// ---- 时间转秒 / Times to seconds ----
tHoldMaxS := TIME_TO_REAL(tHoldMax) / 1000.0;   // 上限秒值 / Hold max [s]
tCycleS   := TIME_TO_REAL(tCycle) / 1000.0;     // 周期秒值 / Cycle [s]

// ---- 启动沿检测（无条件周期刷新）/ Start edge, unconditional refresh ----
rtrigStart(CLK := bSpliceStart);    // 沿检测 / Edge detection

// ---- 非有限与周期合法性闸 / Finite and cycle validity gate ----
IF (tCycle = T#0MS) OR (tCycleS < 0.001) OR (tCycleS > 0.2)
   OR (fTensionA_N <> fTensionA_N) OR (ABS(fTensionA_N) >= 1.0E12)
   OR (fTensionANow_N <> fTensionANow_N) OR (ABS(fTensionANow_N) >= 1.0E12)
   OR (fTensionBSp_N <> fTensionBSp_N) OR (ABS(fTensionBSp_N) >= 1.0E12)
   OR (fRamp_Ns <> fRamp_Ns) OR (ABS(fRamp_Ns) >= 1.0E12)
   OR (fDevMax_N <> fDevMax_N) OR (ABS(fDevMax_N) >= 1.0E12) THEN
    bHoldActive := FALSE;       // 交接退出 / Handover off
    bHoldLatch  := FALSE;       // 锁存复位（本闸自动恢复）/ Latch reset
    eErr := 16#0004_0346;       // 故障码 / Fault code
    RETURN;                     // 给定保持不动 / Command holds
END_IF

// ---- 组态错闸 / Configuration fault gate ----
IF (fRamp_Ns <= 0.0) OR (fTensionBSp_N <= 0.0)
   OR (tHoldMax = T#0MS) OR (tHoldMaxS < 0.1) OR (tHoldMaxS > 30.0) THEN
    bHoldActive := FALSE;       // 交接退出 / Handover off
    eErr := 16#0004_0347;       // 故障码 / Fault code
    RETURN;                     // 本拍结束 / End of cycle
END_IF

// ---- 首扫初始化（R16 纪律：首扫 bCutPermit=FALSE）/ First-scan init ----
IF xFirstScan THEN
    fTensionCmd_N := fTensionANow_N;    // 给定对齐 A 当前指令 / Command aligns to A
    fBlendPct := 0.0;           // B 权重 0 / Blend 0
    bCutPermit := FALSE;        // 裁切禁止 / Cut denied
    bHandoverDone := FALSE;     // 脉冲复位 / Pulse reset
    bHoldActive := FALSE;       // 非交接 / Inactive
    xFirstScan := FALSE;        // 清标记 / Clear flag
END_IF

// ---- 完成脉冲单拍化（上拍 TRUE 本拍清）/ Done pulse: one cycle only ----
IF bHandoverDone THEN
    bHandoverDone := FALSE;     // 下一拍清 / Clear next cycle
END_IF

// ---- 使能撤销 / Disable ----
IF NOT bEnable THEN
    bHoldActive := FALSE;       // 交接退出 / Handover off
    bHoldLatch := FALSE;        // 锁存复位 / Latch reset
    bDevFrozen := FALSE;        // 冻结复位 / Freeze reset
    bCutPermit := FALSE;        // 裁切禁止 / Cut denied
    fBlendPct := 0.0;           // 权重回 0 / Blend 0
    eErr := 16#0004_0345;       // 信息级：未启动 / Info: idle
    RETURN;                     // 本拍结束 / End of cycle
END_IF

// ---- 超时中止锁存与解除 / Abort latch and release ----
IF bHoldLatch THEN
    bHoldActive := FALSE;       // 交接退出 / Handover off
    bCutPermit  := FALSE;       // 绝不裁切 / Never cut
    eErr := 16#0004_0349;       // 故障码回放（给定停在中间值不回退）/ Replay, command holds
    IF bReset THEN
        bHoldLatch := FALSE;    // 解除锁存 / Release latch
        fBlendPct := 0.0;       // 权重回 0 / Blend reset
        fTensionCmd_N := fTensionANow_N;    // 给定对齐 A / Realign to A
    END_IF
    RETURN;                     // 本拍结束 / End of cycle
END_IF

// ---- B 实测无效：拒绝启动（给定不变）/ B invalid: refuse to start ----
IF NOT bBMeasValid THEN
    bHoldActive := FALSE;       // 不启动交接 / Not started
    bCutPermit  := FALSE;       // 裁切禁止 / Cut denied
    eErr := 16#0004_0345;       // 信息级：未启动 / Info: idle
    RETURN;                     // 给定保持不动 / Command holds
END_IF

// ---- 启动沿受理（B 有效才受理）/ Accept start edge with valid B ----
IF rtrigStart.Q AND (fBlendPct < 100.0) AND (NOT bDevFrozen) THEN
    fStartCmd := fTensionCmd_N; // 快照起始给定 / Snapshot start command
    bHoldActive := TRUE;        // 交接进行 / Active
    bDevFrozen := FALSE;        // 冻结复位 / Freeze reset
END_IF

// ---- 单拍给定增量 / Step per cycle ----
fStepN := fRamp_Ns * tCycleS;   // N/s × s = N / Step [N]

// ---- 交接进行路径 / Handover active path ----
IF bHoldActive THEN
    // 交接中张力偏差超限 → 立即冻结斜坡与权重（保张力优先）/ Deviation over limit: freeze
    IF ABS(fTensionA_N - fTensionCmd_N) > fDevMax_N THEN
        bDevFrozen := TRUE;     // 冻结标志 / Freeze flag
        eErr := 16#0004_0348;   // 信息级：冻结 / Info: frozen
    ELSE
        bDevFrozen := FALSE;    // 偏差恢复 → 解除冻结 / Unfreeze
    END_IF

    IF NOT bDevFrozen THEN
        // 分母防护：B 目标与起点重合则直接完成 / Denominator guard: equal targets → done
        IF ABS(fTensionBSp_N - fStartCmd) < 0.001 THEN
            fBlendPct := 100.0;     // 权重直接满 / Blend full
        ELSE
            fBlendPct := fBlendPct + (fStepN / ABS(fTensionBSp_N - fStartCmd)) * 100.0;   // 权重按斜坡推进 / Blend advance
        END_IF
        // 单调递增且钳 [0,100] / Monotonic, clamp
        IF fBlendPct > 100.0 THEN
            fBlendPct := 100.0; // 上限 / Upper clamp
        ELSIF fBlendPct < 0.0 THEN
            fBlendPct := 0.0;   // 下限保护 / Lower guard
        END_IF
        // 给定从 A 起点向 B 目标斜坡过渡 / Command ramps from A start to B target
        fTensionCmd_N := fStartCmd + (fTensionBSp_N - fStartCmd) * fBlendPct / 100.0;   // 插值 / Interpolated
    END_IF

    // ---- 交接完成判 / Completion check ----
    IF fBlendPct >= 100.0 THEN
        fTensionCmd_N := fTensionBSp_N;     // 给定收口到 B 目标 / Command to B target
        fBlendPct := 100.0;     // 权重收口 / Blend full
        bHoldActive := FALSE;   // 交接结束 / Handover off
        bHandoverDone := TRUE;  // 完成脉冲（单拍）/ Done pulse
        eErr := 16#0004_0345;   // 信息级：交接完成 / Info: done
    ELSE
        // ---- 超时监控 / Timeout monitor ----
        tonHold(IN := TRUE, PT := tHoldMax);    // 定时器无条件刷新 / Unconditional refresh
        IF tonHold.Q THEN
            bHoldActive := FALSE;   // 中止交接 / Abort handover
            bHoldLatch := TRUE;     // 锁存 / Latch
            bCutPermit := FALSE;    // 绝不裁切 / Never cut
            eErr := 16#0004_0349;   // 故障码 / Fault code
            RETURN;                 // 本拍结束 / End of cycle
        END_IF
    END_IF
ELSE
    // 非交接期：给定保持，正常码 / Inactive: command holds
    IF eErr <> 16#0004_0348 THEN
        eErr := 16#0004_0345;   // 信息级：未启动 / Info: idle
    END_IF
    tonHold(IN := FALSE, PT := tHoldMax);   // 定时器复位 / Timer reset
END_IF

// ---- 裁切许可：仅权重满且无故障才 TRUE / Cut permit: full blend and no fault ----
bCutPermit := (fBlendPct >= 100.0)
              AND (eErr <> 16#0004_0349)
              AND (eErr <> 16#0004_0347)
              AND (eErr <> 16#0004_0346);   // 许可判 / Permit verdict

END_FUNCTION_BLOCK

(* ---- FB_DL_FilmTaperTension.st ---- *)
(*
  Component : FB_DL_FilmTaperTension
  Category  : DL_Motion
  Type      : FB
  Version   : 1.0.0
  CodeSeg   : 16#04_0_6C
  Summary   : 薄膜锥度张力给定曲线：卷径计算 + 锥度张力给定 + 收卷闭环握手（VAR_IN_OUT）。
              Film taper tension setpoint: roll diameter calculation plus taper curve with a winding handshake via VAR_IN_OUT.
  溯源声明  : 道莅自研 clean-room
  边界安全  : 卷径最小值域闸（> 最小卷径常量，防除零，按派单要点）；膜厚正域闸（> 0）；
              锥度系数为 0 时退化为恒张力（按派单要点）；张力给定钳非负下限；
              与 FB_DL_WindingTensionCtrl 的握手经 VAR_IN_OUT（ioTensionAck），不写其内部状态；
              全浮点比较带 fEps 容差；计数防回卷。
  复用      : 与 FB_DL_WindingTensionCtrl 握手（VAR_IN_OUT 引脚级，无实例依赖）
*)

FUNCTION_BLOCK FB_DL_FilmTaperTension
VAR_INPUT
    bRun        : BOOL;                 (* 给定使能 · Enable *)
    fCoreDiaM   : LREAL := 0.075;       (* 卷芯直径 [m] · Core diameter *)
    fFilmThickUm: LREAL := 20.0;        (* 膜厚 [um] · Film thickness *)
    nTurns      : DINT;                 (* 已卷圈数 [圈] · Wrapped turns *)
    fTensionBaseN: LREAL := 50.0;       (* 外层基准张力 [N] · Base tension at full roll *)
    fTaperK     : LREAL := 0.5;         (* 锥度系数 [比值]，0 为恒张力 · Taper coefficient *)
    fDiaRefM    : LREAL := 0.60;        (* 锥度参考卷径 [m] · Taper reference diameter *)
    fEps        : LREAL := 1.0E-6;      (* 浮点判零容差 [实数域] · Floating zero tolerance *)
END_VAR
VAR_IN_OUT
    ioTensionAck: BOOL;                 (* 收卷闭环握手应答 [引脚]，由张力控件置位 · Handshake ack from the winding ctrl *)
END_VAR
VAR_OUTPUT
    fDiaM       : LREAL;                (* 当前卷径 [m] · Current roll diameter *)
    fTensionSetN: LREAL;                (* 张力给定输出 [N] · Tension setpoint output *)
    bDiaReady   : BOOL;                 (* 卷径有效标志 · Diameter validity flag *)
    bHandshakeOk: BOOL;                 (* 握手应答有效 [开关] · Handshake accepted *)
    bError      : BOOL;                 (* 故障标志，与故障码配对 · Fault flag paired with codes *)
    uErrorId    : UDINT;                (* 事件码 16#0000_006C，0 无事件 · Event code *)
END_VAR
VAR
    uCode   : WORD;     (* 码位暂存，每拍重算 [码] · Code staging *)
    bSigOk  : BOOL;     (* 输入有效标志 · Input validity flag *)
    fDiaMin : LREAL;    (* 最小卷径域值 [m] · Minimum diameter *)
    fRatio  : LREAL;    (* 参考卷径比 [比值] · Diameter ratio *)
    nCycles : UDINT;    (* 有效给定拍计数 [拍]，防回卷 · Valid setpoint count *)
END_VAR
VAR CONSTANT
    DL_FTT_UM2M : LREAL := 1.0E-6;      (* um 到 m 系数 [m/um] · Micrometers to meters *)
    DL_FTT_WRAP : UDINT := 4294967290;  (* 计数防回卷余量 [拍] · Counter wrap guard *)
END_VAR

(* === 段 0 · 实例刷新 === *)
(* 无 TON/R_TRIG 实例：给定按拍直算；No timer instances, direct per-scan setpoint *)

(* === 段 1 · 输入校验与量程闸 === *)
uCode := 16#0000;                       // 每拍清码（可达清零基线）/ Clear codes each scan
fDiaMin := fCoreDiaM + fEps;            (* 最小卷径域值 [m] / Minimum diameter *)
bSigOk := (fCoreDiaM = fCoreDiaM) AND (fFilmThickUm = fFilmThickUm) // 非有限拦截 / Non-finite guard
          AND (fTensionBaseN = fTensionBaseN) AND (fDiaRefM = fDiaRefM)
          AND (ABS(fCoreDiaM) < 1.0E308) AND (ABS(fDiaRefM) < 1.0E308)  // Inf 上限判据 / Inf limits
          AND (fCoreDiaM > fEps)                                        // 卷芯正域闸 / Core diameter gate
          AND (fFilmThickUm > fEps)                                     // 膜厚正域闸 / Thickness gate
          AND (fTensionBaseN >= 0.0)                                    // 张力非负域闸 / Non-negative tension
          AND (fTaperK >= 0.0)                                          // 锥度系数非负闸 / Taper coefficient gate
          AND (fDiaRefM > fEps) AND (nTurns >= 0);                      // 参考卷径/圈数域闸 / Reference and turns gates
IF NOT bSigOk THEN
    uCode := 16#006C;                   // 故障级：域外，给定冻结 / Fault: domain invalid
END_IF

(* === 段 2 · 主逻辑：卷径计算与锥度张力给定 === *)
IF bSigOk THEN
    fDiaM := fCoreDiaM + 2.0 * DINT_TO_LREAL(nTurns) * fFilmThickUm * DL_FTT_UM2M;
                                        (* 卷径 = 芯径 + 2×圈数×膜厚 [m] / Diameter from turns *)
    IF fDiaM < fDiaMin THEN
        fDiaM := fDiaMin;               (* 卷径最小值防御（防除零）/ Minimum diameter guard *)
    END_IF
    bDiaReady := TRUE;                  (* 卷径有效 / Diameter valid *)
    IF fTaperK < fEps THEN
        fTensionSetN := fTensionBaseN;  (* 锥度系数为 0：退化为恒张力 / Zero taper: constant tension *)
    ELSE
        fRatio := fDiaRefM / fDiaM;     (* 参考卷径比（分母已最小值防御）/ Diameter ratio *)
        fTensionSetN := fTensionBaseN * (1.0 + fTaperK * (fRatio - 1.0));
                                        (* 锥度张力给定 [N]：内层紧外层松 / Taper tension setpoint *)
        IF fTensionSetN < 0.0 THEN
            fTensionSetN := 0.0;        (* 给定钳非负下限 / Clamp non-negative *)
        END_IF
    END_IF
END_IF

(* === 段 3 · 输出映射与故障码 === *)
bHandshakeOk := ioTensionAck;           (* 握手应答直读映射（引脚级，不写对方内部）/ Handshake mapping *)
IF bSigOk THEN
    IF nCycles < DL_FTT_WRAP THEN
        nCycles := nCycles + 1;         (* 有效给定计数 / Count valid setpoints *)
    END_IF
END_IF
bError := (uCode <> 16#0000);           (* 故障标志配对 / Fault flag paired *)
uErrorId := WORD_TO_UDINT(uCode);       (* 码位单点写入（16#0000_006C 形态）/ Single write point *)
END_FUNCTION_BLOCK

(* ---- FB_DL_FilmTensionStepper.st ---- *)
(*
  FB_DL_FilmTensionStepper  —  收卷步进张力叠加微调 / Rewinder stepped tension overlay trim
  分类 Category : DL_Motion
  码位 Code     : 16#04_0_A0
  版本 Version  : 1.0.0
  溯源 Source   : LGF Technology 语义借鉴 · clean-room 实现，仅借分类/参数域/命名，未复制源码
  功能 Function : 1) 张力偏差经限斜率步进累加为叠加偏置，叠加量限幅到张力带允许域（防累计漂移把轴拉飞）；
                  2) 只在叠加通道写入，不改基础轴目标（叠加 != 改目标）；
                  3) 张力反馈无效时冻结叠加并保持末次有效偏置，恢复后从保持点继续（无扰）。
  边界 Boundary : ① 叠加偏置总量限幅到张力带允许域（±fOffsetMax）；
                  ② 步进增量限斜率（每拍 <= fStepMax），且只写叠加通道不改基础轴目标；
                  ③ 张力反馈无效时冻结叠加并保持末次有效偏置；
                  ④ 输出三行同向：叠加偏置 → 合成位置 → 冻结标志。
  依赖 Depends  : FB_DL_SuperimposedMove（叠加通道执行，每拍无条件调用）

  码表 Error codes（本件子码步进 16#10，避让邻件码位）:
    16#0002_04A0 故障级：组态非法（增益/步进/叠加上限/任务周期 <= 0 或张力带上下限倒置）
    16#0002_04B0 故障级：叠加层执行故障（映射自依赖实例的故障标志）
    16#0002_04C0 信息级：张力反馈无效，叠加已冻结（不置 bError）
*)

TYPE E_DL_FtsPhase :
(
    eIdle    := 0,   // 空闲 / Idle
    eTrim    := 10,  // 叠加微调 / Overlay trimming
    eFrozen  := 20,  // 反馈无效冻结 / Frozen by invalid feedback
    eFault   := 90   // 故障锁定 / Fault locked
);
END_TYPE

FUNCTION_BLOCK FB_DL_FilmTensionStepper
VAR_INPUT
    bEnable       : BOOL;                          // 总使能，FALSE 冻结叠加 / Master enable
    bReset        : BOOL;                          // 复位，上升沿清故障并归零叠加 / Reset, clears fault and zeroes overlay
    bZeroNow      : BOOL;                          // 叠加归零请求（走斜坡）/ Overlay zero request
    fTensionActN  : REAL;                          // 张力实测反馈 [N]，域 > 0 / Measured tension feedback [N]
    fTensionSpN   : REAL := 50.0;                  // 张力设定 [N]，域 > 0 / Tension setpoint [N]
    fBandN        : REAL := 5.0;                   // 张力带半宽 [N]，域 > 0 / Tension band half width [N]
    fOffsetMaxMm  : REAL := 3.0;                   // 叠加偏置上限 [mm]，域 > 0 / Overlay magnitude limit [mm]
    fOffsetSpeed  : REAL := 2.0;                   // 叠加斜坡限速 [mm/s]，域 > 0 / Overlay ramp speed [mm/s]
    fStepMaxMm    : REAL := 0.05;                  // 单拍步进上限 [mm]，域 > 0 / Step limit per scan [mm]
    fGainMmPerN   : REAL := 0.02;                  // 偏差到偏置增益 [mm/N]，域 > 0 / Error-to-offset gain
    fBasePosMm    : REAL := 0.0;                   // 基础轴位置（仅读，不改）/ Base axis position, read only
    fTaskCycle    : REAL := 0.01;                  // 任务周期 [s]，域 > 0 / Task cycle [s]
    fEps          : REAL := 1.0E-6;                // 浮点判零容差 [1] / Floating zero tolerance
END_VAR
VAR_OUTPUT
    fOffsetCmdMm  : REAL;                          // 叠加偏置指令 [mm]（仅叠加通道）/ Overlay offset command [mm]
    fOffsetActMm  : REAL;                          // 叠加偏置实际值 [mm] / Actual overlay offset [mm]
    fSuperPosMm   : REAL;                          // 合成位置 [mm] = 基础 + 叠加 / Superimposed position [mm]
    bLimited      : BOOL;                          // 偏置已限幅标志 / Offset limited flag
    bFrozen       : BOOL;                          // 叠加冻结标志（保持型）/ Overlay frozen, held
    bError        : BOOL;                          // 故障标志，与故障级码配对 / Fault flag paired with fault codes
    uErrorId      : UDINT;                         // 事件码，0 = 无事件 / Event code, 0 = none
    eStateOut     : E_DL_FtsPhase;                 // 状态机当前态，段尾单点映射 / Phase mapped at tail
END_VAR
VAR
    _eState       : E_DL_FtsPhase := E_DL_FtsPhase.eIdle;  // 内部状态 / Internal state
    rtrReset      : R_TRIG;                        // 复位沿 / Reset edge
    fbOverlay     : FB_DL_SuperimposedMove;        // 叠加通道实例（无条件调用）/ Superimposed move instance
    bCfgOk        : BOOL;                          // 组态合法标志 / Configuration valid
    bFbOk         : BOOL;                          // 张力反馈有效 / Feedback valid
    bInBand       : BOOL;                          // 偏差在张力带内（含容差）/ Error inside band
    fErrN         : REAL;                          // 张力偏差 [N] = 设定 − 实测 / Tension error [N]
    fStepMm       : REAL;                          // 本拍步进量 [mm] / Step this scan [mm]
    fCmdNextMm    : REAL;                          // 下一拍偏置指令 [mm] / Next offset command [mm]
    fCmdHoldMm    : REAL;                          // 保持的偏置指令 [mm] / Held offset command [mm]
    uFault        : UDINT;                         // 锁存故障码 / Latched fault code
    uInfo         : UDINT;                         // 信息级码 / Information code
END_VAR
VAR CONSTANT
    DL_FTS_TMAX   : REAL := 10000.0;               // 张力物理域上限 [N] / Tension domain high [N]
    DL_FTS_MMMAX  : REAL := 100.0;                 // 偏置物理域上限 [mm] / Offset domain high [mm]
END_VAR

(* === 段 0 · 实例刷新（无条件周期调用）=== *)
rtrReset(CLK := bReset);                          // 每拍刷新复位沿

(* === 段 1 · 组态闸与反馈域闸 === *)
bCfgOk := (fGainMmPerN > fEps) AND (fStepMaxMm > fEps) AND (fOffsetMaxMm > fEps)
          AND (fOffsetSpeed > fEps) AND (fTaskCycle > fEps) AND (fBandN > fEps)
          AND (fTensionSpN > fEps) AND (fOffsetMaxMm <= DL_FTS_MMMAX)
          AND (fGainMmPerN = fGainMmPerN) AND (fTensionSpN = fTensionSpN);   // 含 NaN 自反
IF NOT bCfgOk THEN
    uFault := 16#0002_04A0;                       // 故障级：组态非法
END_IF
IF rtrReset.Q AND bCfgOk THEN
    uFault := 16#0000;                            // 复位沿清锁存（复位路径可达）
    fCmdHoldMm := 0.0;                            // 复位归零偏置
    bFrozen := FALSE;                             // 冻结标志同步复位
END_IF
uInfo := 16#0000;                                 // 信息码每拍清零
bFbOk := (fTensionActN = fTensionActN) AND (ABS(fTensionActN) < 1.0E30)
         AND (fTensionActN > 0.0) AND (fTensionActN <= DL_FTS_TMAX);   // NaN 自反 + 正域闸
IF bFbOk THEN
    fErrN := fTensionSpN - fTensionActN;          // 偏差 = 设定 − 实测
    bInBand := ABS(fErrN) <= (fBandN + fEps);     // 带内判据（浮点容差）
ELSE
    fErrN := 0.0;                                 // 无效反馈：偏差不出结论
    bInBand := TRUE;                              // 无效时视作带内（不动叠加）
END_IF

(* === 段 2 · 主状态机（ENUM + CASE，含 ELSE 兜底）=== *)
CASE _eState OF
E_DL_FtsPhase.eIdle :
    fCmdNextMm := fCmdHoldMm;                     // 空闲保持当前偏置
    IF uFault <> 16#0000 THEN
        _eState := E_DL_FtsPhase.eFault;          // 故障优先
    ELSIF NOT bEnable THEN
        _eState := E_DL_FtsPhase.eFrozen;         // 失能即冻结
    ELSIF NOT bFbOk THEN
        bFrozen := TRUE;                          // 反馈无效：冻结
        uInfo := 16#0002_04C0;                    // 信息级：叠加已冻结
        _eState := E_DL_FtsPhase.eFrozen;
    ELSIF bEnable THEN
        _eState := E_DL_FtsPhase.eTrim;           // 进入微调相
    END_IF

E_DL_FtsPhase.eTrim :
    bFrozen := FALSE;                             // 微调相不冻结
    IF (NOT bEnable) OR (NOT bFbOk) THEN
        bFrozen := TRUE;                          // 反馈丢失/失能：冻结
        uInfo := 16#0002_04C0;                    // 信息级：叠加已冻结
        _eState := E_DL_FtsPhase.eFrozen;
    ELSIF bInBand THEN
        fCmdNextMm := fCmdHoldMm;                 // 带内：保持偏置（不继续累加）
        IF bZeroNow THEN
            fCmdNextMm := 0.0;                    // 归零请求：目标置 0（仍走斜坡）
        END_IF
    ELSE
        fStepMm := fErrN * fGainMmPerN;           // 偏差折算步进
        IF fStepMm > fStepMaxMm THEN
            fStepMm := fStepMaxMm;                // 步进上限（正向限斜率）
        END_IF
        IF fStepMm < -fStepMaxMm THEN
            fStepMm := -fStepMaxMm;               // 步进下限（负向限斜率）
        END_IF
        fCmdNextMm := fCmdHoldMm + fStepMm;       // 累加步进
        IF fCmdNextMm > fOffsetMaxMm THEN
            fCmdNextMm := fOffsetMaxMm;           // 叠加总量上限（防漂移拉飞）
        END_IF
        IF fCmdNextMm < -fOffsetMaxMm THEN
            fCmdNextMm := -fOffsetMaxMm;          // 叠加总量下限
        END_IF
    END_IF
    fCmdHoldMm := fCmdNextMm;                     // 偏置指令记账（仅叠加通道）
    IF ABS(fCmdNextMm) >= (fOffsetMaxMm - fEps) THEN
        bLimited := TRUE;                         // 触限标志
    ELSE
        bLimited := FALSE;                        // 未触限，逐拍重算
    END_IF

E_DL_FtsPhase.eFrozen :
    bFrozen := TRUE;                              // 冻结标志保持
    fCmdNextMm := fCmdHoldMm;                     // 保持末次有效偏置（不清零、不外推）
    IF bFbOk AND bEnable AND (uFault = 16#0000) THEN
        bFrozen := FALSE;                         // 反馈恢复：解冻（可到达的解除路径）
        uInfo := 16#0000;                         // 信息码清除
        _eState := E_DL_FtsPhase.eTrim;           // 从保持点继续（无扰）
    END_IF

E_DL_FtsPhase.eFault :
    bFrozen := TRUE;                              // 故障态冻结
    fCmdNextMm := fCmdHoldMm;                     // 保持偏置（不追发新指令）
    IF uFault = 16#0000 THEN
        _eState := E_DL_FtsPhase.eIdle;           // 解锁回空闲
    END_IF

ELSE
    _eState := E_DL_FtsPhase.eFault;              // 非法状态拦截
    uFault := 16#0002_04A0;                       // 故障级：相 ID 越界
    bFrozen := TRUE;                              // 安全侧冻结
    fCmdNextMm := 0.0;                            // 安全侧偏置 0
END_CASE

(* === 段 3 · 叠加通道实例（每拍无条件调用，只写叠加不改基础目标）=== *)
fbOverlay(bEnable := bEnable AND (NOT bFrozen) AND (uFault = 16#0000),   // 冻结/故障时不推进斜坡
          fBasePos := fBasePosMm,                 // 基础轴位置（只读，不改目标）
          fOffsetCmd := fCmdNextMm,               // 叠加偏置指令
          fMaxOffset := fOffsetMaxMm,             // 偏移限幅
          fMaxOffsetSpeed := fOffsetSpeed,        // 偏移斜坡限速
          fTaskCycle := fTaskCycle,               // 任务周期
          bZeroNow := bZeroNow AND (NOT bFrozen));// 归零请求（冻结期间不生效）

(* === 段 4 · 输出映射（三行同向：偏置 → 合成位置 → 冻结标志）=== *)
fOffsetCmdMm := fCmdNextMm;                       // 偏置指令输出
IF fbOverlay.bActive THEN
    fOffsetActMm := fbOverlay.fOffsetAct;         // 叠加实际值
    fSuperPosMm := fbOverlay.fSuperPos;           // 合成位置
ELSE
    fOffsetActMm := fCmdHoldMm;                   // 未激活：保持偏置
    fSuperPosMm := fBasePosMm + fCmdHoldMm;       // 合成位置按记账值计算
END_IF
IF fbOverlay.bError THEN
    uFault := 16#0002_04B0;                       // 故障级：叠加层执行故障（映射依赖实例）
END_IF
bError := (uFault <> 16#0000);                    // 故障标志仅由故障级码置位（R45 配对）
IF bError THEN
    uErrorId := uFault;                           // 故障级优先上报
ELSE
    uErrorId := uInfo;                            // 否则上报信息级码
END_IF
eStateOut := _eState;                             // 输出枚举段尾单点映射（N2 规则）
END_FUNCTION_BLOCK
